// TwinCAT 3 PLC project TcoIo
// Title: TcoIo
// Company: Vortex.Library
// Author: Inxton
// ProjectVersion: 0.6.0.913
// ProgramVersion: 3.1.4023.0
// libraries:
//   Tc2_EtherCAT, * (Beckhoff Automation GmbH)
//   Tc2_Standard, * (Beckhoff Automation GmbH)
//   Tc2_System, * (Beckhoff Automation GmbH)
//   Tc3_Module, * (Beckhoff Automation GmbH)
//   TcoCore, 0.6.0.913 (Vortex.Library)
// project tree:
//   Diagnostics/EtherCAT/MasterDevice/Base/ EtcMasterBase_62654B43.TcDUT, SyncUnitsBase_AD6C35CE.TcDUT, SyncUnitTaskBase_FCD3CBF3.TcDUT, SyncUnitTasksBase_7C8711EB.TcDUT
//   Diagnostics/EtherCAT/MasterDevice/SyncUnit/ InfoData_8649EEEB.TcDUT, ITcoSyncUnit.TcIO, SyncUnitState.TcDUT, SyncUnitTask_AB2F5079.TcDUT, TcoSyncUnit.TcPOU
//   Diagnostics/EtherCAT/SlaveDevice/Base/ EtcSlaveBase_82538BE2.TcDUT, EtcSlaveBoxBase_77A0E4A7.TcDUT, EtcSlaveEndTerminalBase_866C7F0C.TcDUT, EtcSlaveTerminalBase_947E5A46.TcDUT
//   Diagnostics/EtherCAT/MasterDevice/ InfoData_84133AC9.TcDUT, Inputs_A65FACA4.TcDUT, Outputs_23C0ED1D.TcDUT, TcoEthercatDiagnosticsTask.TcPOU, TcoEthercatMasterDeviceState.TcDUT, ITcoEthercatMasterDevice.TcIO, TcoEthercatMasterDevice.TcPOU
//   Diagnostics/EtherCAT/MasterDevice/Messenger/ DiagnosticsMessenger.TcPOU, DiagnosticsMessengers.TcPOU
//   Diagnostics/EtherCAT/SlaveDevice/InfoData/ InfoData_23CBA837.TcDUT, InfoData_6F19DB2B.TcDUT
//   Diagnostics/EtherCAT/SlaveDevice/Inputs/ InputBase_8311D824.TcDUT
//   Diagnostics/EtherCAT/SlaveDevice/Outputs/ OutputBase_10CEE7DE.TcDUT
//   Diagnostics/EtherCAT/SlaveDevice/WcState/ WcState_0B2B16F9.TcDUT, WcState_9091E0EB.TcDUT
//   Diagnostics/EtherCAT/ TcoEthercat.TcGVL
//   Diagnostics/ProfinetComponent/ TcoPnIoComponent.TcPOU
//   EtherCAT/ eEcatState.TcDUT, eLinkState.TcDUT, ITcoEcatComponent.TcIO, TcoEcatSlaveState.TcPOU, TcoEcatComponent.TcPOU
//   / PlcTask.TcTTO
//   POUs/ MAIN.TcPOU
//   SpecialPlcTypes/ TcoAmsAddr.TcDUT, TcoAmsNetId.TcDUT
// real-time tasks:
//   TASK PlcTask: cycle T#15ms, priority 12, ADS port 350
//   TASK PlcTask1: cycle T#15ms, priority 6, ADS port 351
//   TASK PlcTask2: cycle T#10ms, priority 20, ADS port 352
// I/O:
//   DEVICE Device 1 (EtherCAT) (disabled), AmsNetId 172.20.10.110.2.1
//     Term 1 (EK1200) [EK1200-5000 EtherCAT Power supply (2A E-Bus)]
//       Term 2 (EL6002) [EL6002 Interface 2Ch. (RS232)]
//       Term 3 (EL1809) [EL1809 16Ch. Dig. Input 24V, 3ms]
//       Term 4 (EL2809) [EL2809 16Ch. Dig. Output 24V, 0.5A]
//       Term 5 (EL4004) [EL4004 4Ch. Ana. Output 0-10V, 12bit]
//       Term 6 (EL2809) [EL2809 16Ch. Dig. Output 24V, 0.5A]
//       Term 7 (EL6001) [EL6001 Interface (RS232)]
//       Term 8 (EL9011) [EL9011 End Terminal]
//   DEVICE Device 2 (EtherCAT) (disabled), AmsNetId 172.20.10.110.3.1
//     Term 9 (EK1100) [EK1100 EtherCAT Coupler (2A E-Bus)]
//       Term 10 (EK1122) [EK1122 2 port EtherCAT junction]
//         Term 11 (EK1100) [EK1100 EtherCAT Coupler (2A E-Bus)]
//           Term 12 (EL3174-0002) [EL3174-0002 4Ch. Ana. Input +/-10V, +/-20mA 16 Bit, Isolated Channels]
//           Term 13 (EL6001) [EL6001 Interface (RS232)]
//           Term 14 (EL3011) [EL3011 4Ch. Ana. Input 0-20mA DIFF]
//           Term 15 (EL2008) [EL2008 8Ch. Dig. Output 24V, 0.5A]
//           Term 16 (EL2008) [EL2008 8Ch. Dig. Output 24V, 0.5A]
//           Term 17 (EK1110) [EK1110 EtherCAT extension]
//         Term 18 (EK1100) [EK1100 EtherCAT Coupler (2A E-Bus)]
//           Term 19 (EL1809) [EL1809 16Ch. Dig. Input 24V, 3ms]
//           Term 20 (EL2809) [EL2809 16Ch. Dig. Output 24V, 0.5A]
//           Term 21 (EL1809) [EL1809 16Ch. Dig. Input 24V, 3ms]
//           Term 22 (EL3011) [EL3011 4Ch. Ana. Input 0-20mA DIFF]
//           Term 29 (EL9011) [EL9011 End Terminal]
//         Term 23 (EK1100) [EK1100 EtherCAT Coupler (2A E-Bus)]
//           Term 24 (EK1122) [EK1122 2 port EtherCAT junction]
//             Term 25 (EK1100) [EK1100 EtherCAT Coupler (2A E-Bus)]
//               Term 26 (EL1819) [EL1819 16Ch. Dig. Input 24V, 10µs]
//               Term 27 (EL1819) [EL1819 16Ch. Dig. Input 24V, 10µs]
//               Term 30 (EL9011) [EL9011 End Terminal]
//             Term 28 (EK1100) [EK1100 EtherCAT Coupler (2A E-Bus)]
//               Term 29 (EL2788) [EL2788 8Ch. Dig. Output 24V AC/DC, 2A]
//               Term 30 (EL3773) [EL3773 3 Ch. Power Monitoring, Oversample]
//               Term 31 (EL9011) [EL9011 End Terminal]
//           Term 31 (EL3773) [EL3773 3 Ch. Power Monitoring, Oversample]
//           Term 32 (EL2258) [EL2258 8Ch. Dig Output 24V with Multi-Time-Stamp]
//           Term 33 (EL3164) [EL3164 4Ch. Ana. Input 0-10V]
//           Term 32 (EL9011) [EL9011 End Terminal]
//       Term 34 (EL3403) [EL3403 3Ch. Power Measuring]
//       Term 35 (EL6001) [EL6001 Interface (RS232)]
//       Term 36 (EL3024) [EL3024 4Ch. Ana. Input 4-20mA DIFF]
//       Term 33 (EL9011) [EL9011 End Terminal]
//   DEVICE Device 3 (EtherCAT) (disabled), AmsNetId 172.20.10.110.4.1
//     Term 146 (EK1100) [EK1100 EtherCAT Coupler (2A E-Bus)]
//       Term 147 (EK1122) [EK1122 2 port EtherCAT junction]
//         Term 153 (EK1100) [EK1100 EtherCAT Coupler (2A E-Bus)]
//           Term 154 (EK1122) [EK1122 2 port EtherCAT junction]
//             Term 157 (EK1100) [EK1100 EtherCAT Coupler (2A E-Bus)]
//               Term 159 (EL1809) [EL1809 16Ch. Dig. Input 24V, 3ms]
//             Term 158 (EK1100) [EK1100 EtherCAT Coupler (2A E-Bus)]
//               Term 160 (EL1809) [EL1809 16Ch. Dig. Input 24V, 3ms]
//           Term 155 (EL2008) [EL2008 8Ch. Dig. Output 24V, 0.5A]
//           Term 156 (EL2008) [EL2008 8Ch. Dig. Output 24V, 0.5A]
//         Term 178 (EK1100) [EK1100 EtherCAT Coupler (2A E-Bus)]
//           Term 179 (EK1122) [EK1122 2 port EtherCAT junction]
//             Term 180 (EK1100) [EK1100 EtherCAT Coupler (2A E-Bus)]
//               Term 181 (EL1809) [EL1809 16Ch. Dig. Input 24V, 3ms]
//             Term 182 (EK1100) [EK1100 EtherCAT Coupler (2A E-Bus)]
//               Term 183 (EL1809) [EL1809 16Ch. Dig. Input 24V, 3ms]
//           Term 184 (EL2008) [EL2008 8Ch. Dig. Output 24V, 0.5A]
//           Term 185 (EL2008) [EL2008 8Ch. Dig. Output 24V, 0.5A]
//       Term 186 (EK1122) [EK1122 2 port EtherCAT junction]
//         Term 187 (EK1100) [EK1100 EtherCAT Coupler (2A E-Bus)]
//           Term 188 (EK1122) [EK1122 2 port EtherCAT junction]
//             Term 189 (EK1100) [EK1100 EtherCAT Coupler (2A E-Bus)]
//               Term 193 (EL1809) [EL1809 16Ch. Dig. Input 24V, 3ms]
//             Term 194 (EK1100) [EK1100 EtherCAT Coupler (2A E-Bus)]
//               Term 200 (EL1809) [EL1809 16Ch. Dig. Input 24V, 3ms]
//           Term 204 (EL2008) [EL2008 8Ch. Dig. Output 24V, 0.5A]
//           Term 205 (EL2008) [EL2008 8Ch. Dig. Output 24V, 0.5A]
//         Term 207 (EK1100) [EK1100 EtherCAT Coupler (2A E-Bus)]
//           Term 230 (EK1122) [EK1122 2 port EtherCAT junction]
//             Term 231 (EK1100) [EK1100 EtherCAT Coupler (2A E-Bus)]
//               Term 232 (EL1809) [EL1809 16Ch. Dig. Input 24V, 3ms]
//             Term 233 (EK1100) [EK1100 EtherCAT Coupler (2A E-Bus)]
//               Term 234 (EL1809) [EL1809 16Ch. Dig. Input 24V, 3ms]
//           Term 235 (EL2008) [EL2008 8Ch. Dig. Output 24V, 0.5A]
//           Term 236 (EL2008) [EL2008 8Ch. Dig. Output 24V, 0.5A]
//       Term 148 (EL1809) [EL1809 16Ch. Dig. Input 24V, 3ms]
//       Term 149 (EL1809) [EL1809 16Ch. Dig. Input 24V, 3ms]
//       Term 150 (EL1809) [EL1809 16Ch. Dig. Input 24V, 3ms]
//       Term 151 (EL1809) [EL1809 16Ch. Dig. Input 24V, 3ms]
//       Term 152 (EL1809) [EL1809 16Ch. Dig. Input 24V, 3ms]
//       Term 288 (EK1122) [EK1122 2 port EtherCAT junction]
//         Term 289 (EK1100) [EK1100 EtherCAT Coupler (2A E-Bus)]
//           Term 237 (EK1122) [EK1122 2 port EtherCAT junction]
//             Drive 238 (AX5101-0000-0214) [AX5101-0000-0214 EtherCAT Drive (SoE, 1 Ch.)]
//           Term 293 (EL1809) [EL1809 16Ch. Dig. Input 24V, 3ms]
//         Term 294 (EK1100) [EK1100 EtherCAT Coupler (2A E-Bus)]
//           Term 300 (EL1809) [EL1809 16Ch. Dig. Input 24V, 3ms]
//           Term 304 (EL2008) [EL2008 8Ch. Dig. Output 24V, 0.5A]
//           Term 305 (EL2008) [EL2008 8Ch. Dig. Output 24V, 0.5A]
//         Term 307 (EK1100) [EK1100 EtherCAT Coupler (2A E-Bus)]
//           Term 330 (EK1122) [EK1122 2 port EtherCAT junction]
//             Term 331 (EK1100) [EK1100 EtherCAT Coupler (2A E-Bus)]
//               Term 332 (EL1809) [EL1809 16Ch. Dig. Input 24V, 3ms]
//             Term 333 (EK1100) [EK1100 EtherCAT Coupler (2A E-Bus)]
//               Term 334 (EL1809) [EL1809 16Ch. Dig. Input 24V, 3ms]
//           Term 335 (EL2008) [EL2008 8Ch. Dig. Output 24V, 0.5A]
//           Term 336 (EL2008) [EL2008 8Ch. Dig. Output 24V, 0.5A]
//       Term 1158 (EL2008) [EL2008 8Ch. Dig. Output 24V, 0.5A]
//       Term 1159 (EL2008) [EL2008 8Ch. Dig. Output 24V, 0.5A]
//       Term 1160 (EL2008) [EL2008 8Ch. Dig. Output 24V, 0.5A]
//       Term 1161 (EL2008) [EL2008 8Ch. Dig. Output 24V, 0.5A]
//       Term 1162 (EL2008) [EL2008 8Ch. Dig. Output 24V, 0.5A]
//       Term 1163 (EL2008) [EL2008 8Ch. Dig. Output 24V, 0.5A]
//   DEVICE Device 4 (EtherCAT) (disabled), AmsNetId 172.20.10.110.5.1
//     R1 (EK1100) [EK1100 EtherCAT Coupler (2A E-Bus)]
//       R1_A2_EC (EK1122) [EK1122 2 port EtherCAT junction]
//         Servo_A10_1 (AX5106-0000-0203) [AX5106-0000-0203 EtherCAT Drive (SoE, 1 Ch.)]
//         Servo_A10_2 (AX5106-0000-0203) [AX5106-0000-0203 EtherCAT Drive (SoE, 1 Ch.)]
//         Servo_A10_3 (AX5106-0000-0203) [AX5106-0000-0203 EtherCAT Drive (SoE, 1 Ch.)]
//       R1_A3_EC (EK1122) [EK1122 2 port EtherCAT junction]
//         VI-2 (AES-D-BC-ECAT) [AES Fieldbus Coupler]
//           modules: Module 1 (32 Byte Valve Unit (0x7F))
//         VI-4 (AES-D-BC-ECAT) [AES Fieldbus Coupler]
//           modules: Module 1 (32 Byte Valve Unit (0x7F))
//       R1_A4_EC (EK1122) [EK1122 2 port EtherCAT junction]
//         R1_A4_X1 (EK1100) [EK1100 EtherCAT Coupler (2A E-Bus)]
//           R1_A4_X1_PN (EL6631) [EL6631 PROFINET IO Controller]
//           R1_A4_X1_IA1 (EL1809) [EL1809 16Ch. Dig. Input 24V, 3ms]
//           R1_A4_X1_IA2 (EL1809) [EL1809 16Ch. Dig. Input 24V, 3ms]
//           R1_A4_X1_IA3 (EL1809) [EL1809 16Ch. Dig. Input 24V, 3ms]
//           R1_A4_X1_IA4 (EL1809) [EL1809 16Ch. Dig. Input 24V, 3ms]
//           R1_A4_X1_QA1 (EL2809) [EL2809 16Ch. Dig. Output 24V, 0.5A]
//           R1_A4_X1_QA2 (EL2809) [EL2809 16Ch. Dig. Output 24V, 0.5A]
//           R1_A4_X1_QA3 (EL2809) [EL2809 16Ch. Dig. Output 24V, 0.5A]
//           R1_A4_X1_EndTerminal (EL9010) [EL9010 End Terminal]
//         R1_A4_X2 (EK1100) [EK1100 EtherCAT Coupler (2A E-Bus)]
//           R1_A4_X2_A2 (EK1122) [EK1122 2 port EtherCAT junction]
//             R1_A4_X2_A2_VI1 (AES-D-BC-ECAT) [AES Fieldbus Coupler]
//               modules: Module 1 (32 Byte Valve Unit (0x7F))
//             REX_350 (IMecat) [IMecat]
//           R1_A4_X2_IA1 (EL1809) [EL1809 16Ch. Dig. Input 24V, 3ms]
//           R1_A4_X2_IA2 (EL1809) [EL1809 16Ch. Dig. Input 24V, 3ms]
//           R1_A4_X2_IA3 (EL1809) [EL1809 16Ch. Dig. Input 24V, 3ms]
//           R1_A4_X2_IA4 (EL1809) [EL1809 16Ch. Dig. Input 24V, 3ms]
//           R1_A4_X2_IA5 (EL1809) [EL1809 16Ch. Dig. Input 24V, 3ms]
//           R1_A4_X2_QA1 (EL2809) [EL2809 16Ch. Dig. Output 24V, 0.5A]
//           R1_A4_X2_QA2 (EL2809) [EL2809 16Ch. Dig. Output 24V, 0.5A]
//           R1_A4_X2_QA3 (EL2809) [EL2809 16Ch. Dig. Output 24V, 0.5A]
//           R1_A4_X2_EndTerminal (EL9010) [EL9010 End Terminal]
//       R1_A5_DI (EL1809) [EL1809 16Ch. Dig. Input 24V, 3ms]
//       R1_A6_DI (EL1809) [EL1809 16Ch. Dig. Input 24V, 3ms]
//       R1_A7_DI (EL1809) [EL1809 16Ch. Dig. Input 24V, 3ms]
//       R1_A8_DI (EL1809) [EL1809 16Ch. Dig. Input 24V, 3ms]
//       R1_A9_DI (EL1809) [EL1809 16Ch. Dig. Input 24V, 3ms]
//       R1_A10_DI (EL1809) [EL1809 16Ch. Dig. Input 24V, 3ms]
//       R1_A11_DI (EL1809) [EL1809 16Ch. Dig. Input 24V, 3ms]
//       R1_A12_DI (EL1809) [EL1809 16Ch. Dig. Input 24V, 3ms]
//       R1_A13_DI (EL1809) [EL1809 16Ch. Dig. Input 24V, 3ms]
//       R1_A14_DI (EL1809) [EL1809 16Ch. Dig. Input 24V, 3ms]
//       R1_A15_DI (EL1809) [EL1809 16Ch. Dig. Input 24V, 3ms]
//       R1_A16_DI (EL1809) [EL1809 16Ch. Dig. Input 24V, 3ms]
//       R1_A17_DI (EL1809) [EL1809 16Ch. Dig. Input 24V, 3ms]
//       R1_A18_DO (EL2809) [EL2809 16Ch. Dig. Output 24V, 0.5A]
//       R1_A19_DO (EL2809) [EL2809 16Ch. Dig. Output 24V, 0.5A]
//       R1_A20_DO (EL2809) [EL2809 16Ch. Dig. Output 24V, 0.5A]
//       R1_A21_DO (EL2809) [EL2809 16Ch. Dig. Output 24V, 0.5A]
//       R1_A22_DO (EL2809) [EL2809 16Ch. Dig. Output 24V, 0.5A]
//       R1_A23_DO (EL2809) [EL2809 16Ch. Dig. Output 24V, 0.5A]
//       R1_EndTerminal (EL9011) [EL9011 End Terminal]
//     R2 (EK1100) [EK1100 EtherCAT Coupler (2A E-Bus)]
//       R2_A2_EC (EK1122) [EK1122 2 port EtherCAT junction]
//         Servo_A20-2 (AX5103-0000-0203) [AX5103-0000-0203 EtherCAT Drive (SoE, 1 Ch.)]
//         VI-3 (AES-D-BC-ECAT) [AES Fieldbus Coupler]
//           modules: Module 1 (32 Byte Valve Unit (0x7F))
//       R2_A3_DI (EL1809) [EL1809 16Ch. Dig. Input 24V, 3ms]
//       R2_A4_DI (EL1809) [EL1809 16Ch. Dig. Input 24V, 3ms]
//       R2_A5_DI (EL1809) [EL1809 16Ch. Dig. Input 24V, 3ms]
//       R2_A6_DI (EL1809) [EL1809 16Ch. Dig. Input 24V, 3ms]
//       R2_A7_DI (EL1809) [EL1809 16Ch. Dig. Input 24V, 3ms]
//       R2_A8_DI (EL1809) [EL1809 16Ch. Dig. Input 24V, 3ms]
//       R2_A9_DI (EL1809) [EL1809 16Ch. Dig. Input 24V, 3ms]
//       R2_A10_DI (EL1809) [EL1809 16Ch. Dig. Input 24V, 3ms]
//       R2_A11_DC (EL7332) [EL7332 2Ch. DC motor output stage (24V, 1.5A)]
//       R2_A12_DI (EL1809) [EL1809 16Ch. Dig. Input 24V, 3ms]
//       R2_A13_DI (EL1809) [EL1809 16Ch. Dig. Input 24V, 3ms]
//       R2_A14_DI (EL1809) [EL1809 16Ch. Dig. Input 24V, 3ms]
//       R2_A15_DO (EL2809) [EL2809 16Ch. Dig. Output 24V, 0.5A]
//       R2_A16_DO (EL2809) [EL2809 16Ch. Dig. Output 24V, 0.5A]
//       R2_A17_DO (EL2809) [EL2809 16Ch. Dig. Output 24V, 0.5A]
//       R2_A18_DO (EL2809) [EL2809 16Ch. Dig. Output 24V, 0.5A]
//       R2_A19_DO (EL2809) [EL2809 16Ch. Dig. Output 24V, 0.5A]
//       R2_EndTerminal (EL9011) [EL9011 End Terminal]
//     R3 (EK1100) [EK1100 EtherCAT Coupler (2A E-Bus)]
//       R3_A2_EC (EK1122) [EK1122 2 port EtherCAT junction]
//         R3_FESTO (CMMP-AS V4p0 CiA402) [CMMP-AS V4p0 CiA402]
//         VI-1 (AES-D-BC-ECAT) [AES Fieldbus Coupler]
//           modules: Module 1 (32 Byte Valve Unit (0x7F))
//       R3_A3_DI (EL1809) [EL1809 16Ch. Dig. Input 24V, 3ms]
//       R3_A4_DI (EL1809) [EL1809 16Ch. Dig. Input 24V, 3ms]
//       R3_A5_DI (EL1809) [EL1809 16Ch. Dig. Input 24V, 3ms]
//       R3_A6_DI (EL1809) [EL1809 16Ch. Dig. Input 24V, 3ms]
//       R3_A7_DI (EL1809) [EL1809 16Ch. Dig. Input 24V, 3ms]
//       R3_A8_DI (EL1809) [EL1809 16Ch. Dig. Input 24V, 3ms]
//       R3_A9_DO (EL2809) [EL2809 16Ch. Dig. Output 24V, 0.5A]
//       R3_A10_DO (EL2809) [EL2809 16Ch. Dig. Output 24V, 0.5A]
//       R3_EndTerminal (EL9011) [EL9011 End Terminal]
//     R4 (EK1100) [EK1100 EtherCAT Coupler (2A E-Bus)]
//       R4_A2_EC (EK1122) [EK1122 2 port EtherCAT junction]
//         R4_FESTO (CMMP-AS V4p0 CiA402) [CMMP-AS V4p0 CiA402]
//         RH (EK1100) [EK1100 EtherCAT Coupler (2A E-Bus)]
//           RH_A2 (EK1122) [EK1122 2 port EtherCAT junction]
//             RH_SAFETY (Flexi Gateway GETC1) [FLX0-GETC100]
//             RH_A2_X2 (EK1100) [EK1100 EtherCAT Coupler (2A E-Bus)]
//               RH_A2_X2_A2 (EL7211-0010) [EL7211-0010 1Ch. MDP742 Servo motor output stage with OCT (50V, 4.5A RMS)]
//               RH_A2_X2_A3 (EL1809) [EL1809 16Ch. Dig. Input 24V, 3ms]
//               RH_A2_X2_A4 (EL2809) [EL2809 16Ch. Dig. Output 24V, 0.5A]
//               Term 1057 (EL9011) [EL9011 End Terminal]
//           RH_A3 (EL6631) [EL6631 PROFINET IO Controller]
//           RH_A4 (EL1809) [EL1809 16Ch. Dig. Input 24V, 3ms]
//           RH_A5 (EL1809) [EL1809 16Ch. Dig. Input 24V, 3ms]
//           RH_A6 (EL1809) [EL1809 16Ch. Dig. Input 24V, 3ms]
//           RH_A7 (EL2809) [EL2809 16Ch. Dig. Output 24V, 0.5A]
//           RH_A8 (EL1809) [EL1809 16Ch. Dig. Input 24V, 3ms]
//           RH_A9 (EL2809) [EL2809 16Ch. Dig. Output 24V, 0.5A]
//           RH_A10 (EL2809) [EL2809 16Ch. Dig. Output 24V, 0.5A]
//           RH_A11 (EL2809) [EL2809 16Ch. Dig. Output 24V, 0.5A]
//           RH_EndTerminal (EL9011) [EL9011 End Terminal]
//       R4_A3_DI (EL1809) [EL1809 16Ch. Dig. Input 24V, 3ms]
//       R4_A4_DI (EL1809) [EL1809 16Ch. Dig. Input 24V, 3ms]
//       R4_A5_DI (EL1809) [EL1809 16Ch. Dig. Input 24V, 3ms]
//       R4_A6_DI (EL1809) [EL1809 16Ch. Dig. Input 24V, 3ms]
//       R4_A7_DI (EL1809) [EL1809 16Ch. Dig. Input 24V, 3ms]
//       R4_EndTerminal (EL9011) [EL9011 End Terminal]
//     R4A (EK1100) [EK1100 EtherCAT Coupler (2A E-Bus)]
//       A2 (EK1122) [EK1122 2 port EtherCAT junction]
//         VI-7 (AES-D-BC-ECAT) [AES Fieldbus Coupler]
//           modules: Module 1 (32 Byte Valve Unit (0x7F))
//       A3 (EL1809) [EL1809 16Ch. Dig. Input 24V, 3ms]
//       A4 (EL1809) [EL1809 16Ch. Dig. Input 24V, 3ms]
//       A5 (EL1809) [EL1809 16Ch. Dig. Input 24V, 3ms]
//       A6 (EL1809) [EL1809 16Ch. Dig. Input 24V, 3ms]
//       A7 (EL3692) [EL3692 2Ch. resistance measurement terminal]
//       A8 (EL3692) [EL3692 2Ch. resistance measurement terminal]
//       A9 (EL2008) [EL2008 8Ch. Dig. Output 24V, 0.5A]
//       A10 (EL2008) [EL2008 8Ch. Dig. Output 24V, 0.5A]
//       R4A_EndTerminal (EL9011) [EL9011 End Terminal]
//     R5 (EK1100) [EK1100 EtherCAT Coupler (2A E-Bus)]
//       R5_A2_EC (EK1122) [EK1122 2 port EtherCAT junction]
//         VI-5 (AES-D-BC-ECAT) [AES Fieldbus Coupler]
//           modules: Module 1 (32 Byte Valve Unit (0x7F))
//       R5_A3_DI (EL1809) [EL1809 16Ch. Dig. Input 24V, 3ms]
//       R5_A4_DI (EL1809) [EL1809 16Ch. Dig. Input 24V, 3ms]
//       R5_A5_DO (EL2809) [EL2809 16Ch. Dig. Output 24V, 0.5A]
//       R5_A6_DO (EL2809) [EL2809 16Ch. Dig. Output 24V, 0.5A]
//       R5_EndTerminal (EL9011) [EL9011 End Terminal]
//     R6 (EK1100) [EK1100 EtherCAT Coupler (2A E-Bus)]
//       R6_A2_DI (EL1809) [EL1809 16Ch. Dig. Input 24V, 3ms]
//       R6_A3_DI (EL1809) [EL1809 16Ch. Dig. Input 24V, 3ms]
//       R6_A4_DI (EL1809) [EL1809 16Ch. Dig. Input 24V, 3ms]
//       R6_A5_DI (EL1809) [EL1809 16Ch. Dig. Input 24V, 3ms]
//       R6_A6_DI (EL1809) [EL1809 16Ch. Dig. Input 24V, 3ms]
//       R6_A7_DI (EL1809) [EL1809 16Ch. Dig. Input 24V, 3ms]
//       R6_A8_DI (EL1809) [EL1809 16Ch. Dig. Input 24V, 3ms]
//       R6_A9_DI (EL1809) [EL1809 16Ch. Dig. Input 24V, 3ms]
//       R6_A10_DI (EL1809) [EL1809 16Ch. Dig. Input 24V, 3ms]
//       R6_A11_DI (EL1809) [EL1809 16Ch. Dig. Input 24V, 3ms]
//       R6_A12_DI (EL1809) [EL1809 16Ch. Dig. Input 24V, 3ms]
//       R6_A13_DI (EL1809) [EL1809 16Ch. Dig. Input 24V, 3ms]
//       R6_A14_DI (EL1809) [EL1809 16Ch. Dig. Input 24V, 3ms]
//       R6_A15_DO (EL2809) [EL2809 16Ch. Dig. Output 24V, 0.5A]
//       R6_A16_DO (EL2809) [EL2809 16Ch. Dig. Output 24V, 0.5A]
//       R6_A17_DO (EL2809) [EL2809 16Ch. Dig. Output 24V, 0.5A]
//       R6_A18_DO (EL2809) [EL2809 16Ch. Dig. Output 24V, 0.5A]
//       R6_EndTerminal (EL9011) [EL9011 End Terminal]
//     R7 (EK1100) [EK1100 EtherCAT Coupler (2A E-Bus)]
//       R7_A2_EC (EK1122) [EK1122 2 port EtherCAT junction]
//         VI-6 (AES-D-BC-ECAT) [AES Fieldbus Coupler]
//           modules: Module 1 (32 Byte Valve Unit (0x7F))
//       R7_A3_DI (EL1809) [EL1809 16Ch. Dig. Input 24V, 3ms]
//       R7_A4_DI (EL1809) [EL1809 16Ch. Dig. Input 24V, 3ms]
//       R7_A5_DI (EL1809) [EL1809 16Ch. Dig. Input 24V, 3ms]
//       R7_A6_DI (EL1809) [EL1809 16Ch. Dig. Input 24V, 3ms]
//       R7_A7_DI (EL1809) [EL1809 16Ch. Dig. Input 24V, 3ms]
//       R7_A8_DI (EL1809) [EL1809 16Ch. Dig. Input 24V, 3ms]
//       R7_A9_DI (EL1809) [EL1809 16Ch. Dig. Input 24V, 3ms]
//       R7_A10_DI (EL1809) [EL1809 16Ch. Dig. Input 24V, 3ms]
//       R7_A11_DI (EL1809) [EL1809 16Ch. Dig. Input 24V, 3ms]
//       R7_A12_DI (EL1809) [EL1809 16Ch. Dig. Input 24V, 3ms]
//       R7_A13_DI (EL2809) [EL2809 16Ch. Dig. Output 24V, 0.5A]
//       R7_A14_DI (EL2809) [EL2809 16Ch. Dig. Output 24V, 0.5A]
//       R7_EndTerminal (EL9011) [EL9011 End Terminal]
//     R8 (EK1100) [EK1100 EtherCAT Coupler (2A E-Bus)]
//       R8_A2 (EK1122) [EK1122 2 port EtherCAT junction]
//         R8_AB0 (EPP1322-0001) [EPP1322-0001 3 port EtherCAT P gateway]
//           R8_AB24 (EPP1008-0001) [EPP1008-0001 8 Ch. Dig. Input 24V, 3ms, M8]
//           R8_AB23 (EPP1008-0001) [EPP1008-0001 8 Ch. Dig. Input 24V, 3ms, M8]
//           R8_AB22 (EPP1008-0001) [EPP1008-0001 8 Ch. Dig. Input 24V, 3ms, M8]
//           R8_AB21 (EPP1008-0001) [EPP1008-0001 8 Ch. Dig. Input 24V, 3ms, M8]
//           R8_AB20 (EPP1008-0001) [EPP1008-0001 8 Ch. Dig. Input 24V, 3ms, M8]
//           R8_AB19 (EPP1008-0001) [EPP1008-0001 8 Ch. Dig. Input 24V, 3ms, M8]
//           R8_AB18 (EPP1008-0001) [EPP1008-0001 8 Ch. Dig. Input 24V, 3ms, M8]
//           R8_AB17 (EPP1008-0001) [EPP1008-0001 8 Ch. Dig. Input 24V, 3ms, M8]
//           R8_AB16 (EPP1008-0001) [EPP1008-0001 8 Ch. Dig. Input 24V, 3ms, M8]
//           R8_AB15 (EPP1008-0001) [EPP1008-0001 8 Ch. Dig. Input 24V, 3ms, M8]
//           R8_AB14 (EPP1008-0001) [EPP1008-0001 8 Ch. Dig. Input 24V, 3ms, M8]
//           R8_AB13 (EPP1008-0001) [EPP1008-0001 8 Ch. Dig. Input 24V, 3ms, M8]
//           Box 379 (EPP1332-0001) [EPP1332-0001 3 port EtherCAT P junction, power refreshing]
//           R8_AB12 (EPP1008-0001) [EPP1008-0001 8 Ch. Dig. Input 24V, 3ms, M8]
//           R8_AB11 (EPP1008-0001) [EPP1008-0001 8 Ch. Dig. Input 24V, 3ms, M8]
//           R8_AB10 (EPP1008-0001) [EPP1008-0001 8 Ch. Dig. Input 24V, 3ms, M8]
//           R8_AB9 (EPP1008-0001) [EPP1008-0001 8 Ch. Dig. Input 24V, 3ms, M8]
//           R8_AB8 (EPP1008-0001) [EPP1008-0001 8 Ch. Dig. Input 24V, 3ms, M8]
//           R8_AB7 (EPP1008-0001) [EPP1008-0001 8 Ch. Dig. Input 24V, 3ms, M8]
//           R8_AB6 (EPP1008-0001) [EPP1008-0001 8 Ch. Dig. Input 24V, 3ms, M8]
//           R8_AB5 (EPP1008-0001) [EPP1008-0001 8 Ch. Dig. Input 24V, 3ms, M8]
//           R8_AB4 (EPP1008-0001) [EPP1008-0001 8 Ch. Dig. Input 24V, 3ms, M8]
//           R8_AB3 (EPP1008-0001) [EPP1008-0001 8 Ch. Dig. Input 24V, 3ms, M8]
//           R8_AB2 (EPP1008-0001) [EPP1008-0001 8 Ch. Dig. Input 24V, 3ms, M8]
//           R8_AB1 (EPP1008-0001) [EPP1008-0001 8 Ch. Dig. Input 24V, 3ms, M8]
//       R8_A3 (EK1122) [EK1122 2 port EtherCAT junction]
//         VI-10 (AES-D-BC-ECAT) [AES Fieldbus Coupler]
//           modules: Module 1 (32 Byte Valve Unit (0x7F))
//         VI-9 (AES-D-BC-ECAT) [AES Fieldbus Coupler]
//           modules: Module 1 (32 Byte Valve Unit (0x7F))
//       R8_A5 (EL1809) [EL1809 16Ch. Dig. Input 24V, 3ms]
//       R8_A6 (EL2809) [EL2809 16Ch. Dig. Output 24V, 0.5A]
//       R8_A7 (EL2809) [EL2809 16Ch. Dig. Output 24V, 0.5A]
//       R8_A8 (EK1122) [EK1122 2 port EtherCAT junction]
//         RC10_1 (EK1100) [EK1100 EtherCAT Coupler (2A E-Bus)]
//           RC10_A2 (EK1122) [EK1122 2 port EtherCAT junction]
//             RC10_VI (AES-D-BC-ECAT) [AES Fieldbus Coupler]
//               modules: Module 1 (32 Byte Valve Unit (0x7F))
//             RC10_SAFETY (Flexi Soft EtherCAT Gateway) [Flexi Soft EtherCAT Gateway]
//           RC10_A3 (EK1122) [EK1122 2 port EtherCAT junction]
//             RC10_EPP (EPP1322-0001) [EPP1322-0001 3 port EtherCAT P gateway]
//               RC10_AB1 (EPP1008-0001) [EPP1008-0001 8 Ch. Dig. Input 24V, 3ms, M8]
//               RC10_AB2 (EPP1008-0001) [EPP1008-0001 8 Ch. Dig. Input 24V, 3ms, M8]
//               RC10_AB6 (EPP1008-0001) [EPP1008-0001 8 Ch. Dig. Input 24V, 3ms, M8]
//               RC10_AB3 (EPP1008-0001) [EPP1008-0001 8 Ch. Dig. Input 24V, 3ms, M8]
//               RC10_AB4 (EPP1008-0001) [EPP1008-0001 8 Ch. Dig. Input 24V, 3ms, M8]
//               RC10_AB7 (EPP1008-0001) [EPP1008-0001 8 Ch. Dig. Input 24V, 3ms, M8]
//               RC10_AB9 (EPP1008-0001) [EPP1008-0001 8 Ch. Dig. Input 24V, 3ms, M8]
//               RC10_AB10 (EPP1008-0001) [EPP1008-0001 8 Ch. Dig. Input 24V, 3ms, M8]
//               RC10_AB8 (EPP1008-0001) [EPP1008-0001 8 Ch. Dig. Input 24V, 3ms, M8]
//               RC10_AB5 (EPP1008-0001) [EPP1008-0001 8 Ch. Dig. Input 24V, 3ms, M8]
//           RC10_A5 (EL1809) [EL1809 16Ch. Dig. Input 24V, 3ms]
//           RC10_A6 (EL1809) [EL1809 16Ch. Dig. Input 24V, 3ms]
//           RC10_A7 (EL2809) [EL2809 16Ch. Dig. Output 24V, 0.5A]
//           RC10_A8 (EL2809) [EL2809 16Ch. Dig. Output 24V, 0.5A]
//           RC10_A9 (EL2809) [EL2809 16Ch. Dig. Output 24V, 0.5A]
//           RC10_1_EndTerminal (EL9011) [EL9011 End Terminal]
//         RC10_2 (EK1100) [EK1100 EtherCAT Coupler (2A E-Bus)]
//           RC10_B1 (EL7041-1000) [EL7041-1000 1Ch. Stepper motor output stage (50V, 5A, standard)]
//           RC10_B2 (EL7041-1000) [EL7041-1000 1Ch. Stepper motor output stage (50V, 5A, standard)]
//           RC10_C11 (EL7041-1000) [EL7041-1000 1Ch. Stepper motor output stage (50V, 5A, standard)]
//           RC10_C12 (EL7041-1000) [EL7041-1000 1Ch. Stepper motor output stage (50V, 5A, standard)]
//           RC10_C21 (EL7041-1000) [EL7041-1000 1Ch. Stepper motor output stage (50V, 5A, standard)]
//           RC10_C22 (EL7041-1000) [EL7041-1000 1Ch. Stepper motor output stage (50V, 5A, standard)]
//           RC10_2_EndTerminal (EL9010) [EL9010 End Terminal]
//         RC20_1 (EK1100) [EK1100 EtherCAT Coupler (2A E-Bus)]
//           RC20_A2 (EK1122) [EK1122 2 port EtherCAT junction]
//             RC20_VI (AES-D-BC-ECAT) [AES Fieldbus Coupler]
//               modules: Module 1 (32 Byte Valve Unit (0x7F))
//             RC20_SAFETY (Flexi Soft EtherCAT Gateway) [Flexi Soft EtherCAT Gateway]
//           RC20_A3 (EK1122) [EK1122 2 port EtherCAT junction]
//             RC20_EPP (EPP1322-0001) [EPP1322-0001 3 port EtherCAT P gateway]
//               RC20_AB1 (EPP1008-0001) [EPP1008-0001 8 Ch. Dig. Input 24V, 3ms, M8]
//               RC20_AB2 (EPP1008-0001) [EPP1008-0001 8 Ch. Dig. Input 24V, 3ms, M8]
//               RC20_AB6 (EPP1008-0001) [EPP1008-0001 8 Ch. Dig. Input 24V, 3ms, M8]
//               RC20_AB3 (EPP1008-0001) [EPP1008-0001 8 Ch. Dig. Input 24V, 3ms, M8]
//               RC20_AB4 (EPP1008-0001) [EPP1008-0001 8 Ch. Dig. Input 24V, 3ms, M8]
//               RC20_AB7 (EPP1008-0001) [EPP1008-0001 8 Ch. Dig. Input 24V, 3ms, M8]
//               RC20_AB9 (EPP1008-0001) [EPP1008-0001 8 Ch. Dig. Input 24V, 3ms, M8]
//               RC20_AB10 (EPP1008-0001) [EPP1008-0001 8 Ch. Dig. Input 24V, 3ms, M8]
//               RC20_AB8 (EPP1008-0001) [EPP1008-0001 8 Ch. Dig. Input 24V, 3ms, M8]
//               RC20_AB5 (EPP1008-0001) [EPP1008-0001 8 Ch. Dig. Input 24V, 3ms, M8]
//           RC20_A5 (EL1809) [EL1809 16Ch. Dig. Input 24V, 3ms]
//           RC20_A6 (EL1809) [EL1809 16Ch. Dig. Input 24V, 3ms]
//           RC20_A7 (EL2809) [EL2809 16Ch. Dig. Output 24V, 0.5A]
//           RC20_A8 (EL2809) [EL2809 16Ch. Dig. Output 24V, 0.5A]
//           RC20_A9 (EL2809) [EL2809 16Ch. Dig. Output 24V, 0.5A]
//           RC20_1_EndTerminal (EL9010) [EL9010 End Terminal]
//         RC20_2 (EK1100) [EK1100 EtherCAT Coupler (2A E-Bus)]
//           RC20_B1 (EL7041-1000) [EL7041-1000 1Ch. Stepper motor output stage (50V, 5A, standard)]
//           RC20_B2 (EL7041-1000) [EL7041-1000 1Ch. Stepper motor output stage (50V, 5A, standard)]
//           RC20_C11 (EL7041-1000) [EL7041-1000 1Ch. Stepper motor output stage (50V, 5A, standard)]
//           RC20_C12 (EL7041-1000) [EL7041-1000 1Ch. Stepper motor output stage (50V, 5A, standard)]
//           RC20_C21 (EL7041-1000) [EL7041-1000 1Ch. Stepper motor output stage (50V, 5A, standard)]
//           RC20_C22 (EL7041-1000) [EL7041-1000 1Ch. Stepper motor output stage (50V, 5A, standard)]
//           RC20_2_EndTerminal (EL9010) [EL9010 End Terminal]
//       R8_A9 (EK1122) [EK1122 2 port EtherCAT junction]
//         RC30_1 (EK1100) [EK1100 EtherCAT Coupler (2A E-Bus)]
//           RC30_A2 (EK1122) [EK1122 2 port EtherCAT junction]
//             RC30_VI (AES-D-BC-ECAT) [AES Fieldbus Coupler]
//               modules: Module 1 (32 Byte Valve Unit (0x7F))
//             RC30_SAFETY (Flexi Soft EtherCAT Gateway) [Flexi Soft EtherCAT Gateway]
//           RC30_A3 (EK1122) [EK1122 2 port EtherCAT junction]
//             RC30_EPP (EPP1322-0001) [EPP1322-0001 3 port EtherCAT P gateway]
//               RC30_AB1 (EPP1008-0001) [EPP1008-0001 8 Ch. Dig. Input 24V, 3ms, M8]
//               RC30_AB2 (EPP1008-0001) [EPP1008-0001 8 Ch. Dig. Input 24V, 3ms, M8]
//               RC30_AB6 (EPP1008-0001) [EPP1008-0001 8 Ch. Dig. Input 24V, 3ms, M8]
//               RC30_AB3 (EPP1008-0001) [EPP1008-0001 8 Ch. Dig. Input 24V, 3ms, M8]
//               RC30_AB4 (EPP1008-0001) [EPP1008-0001 8 Ch. Dig. Input 24V, 3ms, M8]
//               RC30_AB7 (EPP1008-0001) [EPP1008-0001 8 Ch. Dig. Input 24V, 3ms, M8]
//               RC30_AB9 (EPP1008-0001) [EPP1008-0001 8 Ch. Dig. Input 24V, 3ms, M8]
//               RC30_AB10 (EPP1008-0001) [EPP1008-0001 8 Ch. Dig. Input 24V, 3ms, M8]
//               RC30_AB8 (EPP1008-0001) [EPP1008-0001 8 Ch. Dig. Input 24V, 3ms, M8]
//               RC30_AB5 (EPP1008-0001) [EPP1008-0001 8 Ch. Dig. Input 24V, 3ms, M8]
//           RC30_A5 (EL1809) [EL1809 16Ch. Dig. Input 24V, 3ms]
//           RC30_A6 (EL1809) [EL1809 16Ch. Dig. Input 24V, 3ms]
//           RC30_A7 (EL2809) [EL2809 16Ch. Dig. Output 24V, 0.5A]
//           RC30_A8 (EL2809) [EL2809 16Ch. Dig. Output 24V, 0.5A]
//           RC30_A9 (EL2809) [EL2809 16Ch. Dig. Output 24V, 0.5A]
//           RC30_1_EndTerminal (EL9010) [EL9010 End Terminal]
//         RC30_2 (EK1100) [EK1100 EtherCAT Coupler (2A E-Bus)]
//           RC30_B1 (EL7041-1000) [EL7041-1000 1Ch. Stepper motor output stage (50V, 5A, standard)]
//           RC30_B2 (EL7041-1000) [EL7041-1000 1Ch. Stepper motor output stage (50V, 5A, standard)]
//           RC30_C11 (EL7041-1000) [EL7041-1000 1Ch. Stepper motor output stage (50V, 5A, standard)]
//           RC30_C12 (EL7041-1000) [EL7041-1000 1Ch. Stepper motor output stage (50V, 5A, standard)]
//           RC30_C21 (EL7041-1000) [EL7041-1000 1Ch. Stepper motor output stage (50V, 5A, standard)]
//           RC30_C22 (EL7041-1000) [EL7041-1000 1Ch. Stepper motor output stage (50V, 5A, standard)]
//           RC30_2_EndTerminal (EL9010) [EL9010 End Terminal]
//         RC40_1 (EK1100) [EK1100 EtherCAT Coupler (2A E-Bus)]
//           RC40_A2 (EK1122) [EK1122 2 port EtherCAT junction]
//             RC40_VI (AES-D-BC-ECAT) [AES Fieldbus Coupler]
//               modules: Module 1 (32 Byte Valve Unit (0x7F))
//             RC40_SAFETY (Flexi Soft EtherCAT Gateway) [Flexi Soft EtherCAT Gateway]
//           RC40_A3 (EK1122) [EK1122 2 port EtherCAT junction]
//             RC40_EPP (EPP1322-0001) [EPP1322-0001 3 port EtherCAT P gateway]
//               RC40_AB1 (EPP1008-0001) [EPP1008-0001 8 Ch. Dig. Input 24V, 3ms, M8]
//               RC40_AB2 (EPP1008-0001) [EPP1008-0001 8 Ch. Dig. Input 24V, 3ms, M8]
//               RC40_AB6 (EPP1008-0001) [EPP1008-0001 8 Ch. Dig. Input 24V, 3ms, M8]
//               RC40_AB3 (EPP1008-0001) [EPP1008-0001 8 Ch. Dig. Input 24V, 3ms, M8]
//               RC40_AB4 (EPP1008-0001) [EPP1008-0001 8 Ch. Dig. Input 24V, 3ms, M8]
//               RC40_AB7 (EPP1008-0001) [EPP1008-0001 8 Ch. Dig. Input 24V, 3ms, M8]
//               RC40_AB9 (EPP1008-0001) [EPP1008-0001 8 Ch. Dig. Input 24V, 3ms, M8]
//               RC40_AB10 (EPP1008-0001) [EPP1008-0001 8 Ch. Dig. Input 24V, 3ms, M8]
//               RC40_AB8 (EPP1008-0001) [EPP1008-0001 8 Ch. Dig. Input 24V, 3ms, M8]
//               RC40_AB5 (EPP1008-0001) [EPP1008-0001 8 Ch. Dig. Input 24V, 3ms, M8]
//           RC40_A5 (EL1809) [EL1809 16Ch. Dig. Input 24V, 3ms]
//           RC40_A6 (EL1809) [EL1809 16Ch. Dig. Input 24V, 3ms]
//           RC40_A7 (EL2809) [EL2809 16Ch. Dig. Output 24V, 0.5A]
//           RC40_A8 (EL2809) [EL2809 16Ch. Dig. Output 24V, 0.5A]
//           RC40_A9 (EL2809) [EL2809 16Ch. Dig. Output 24V, 0.5A]
//           RC40_1_EndTerminal (EL9010) [EL9010 End Terminal]
//         RC40_2 (EK1100) [EK1100 EtherCAT Coupler (2A E-Bus)]
//           RC40_B1 (EL7041-1000) [EL7041-1000 1Ch. Stepper motor output stage (50V, 5A, standard)]
//           RC40_B2 (EL7041-1000) [EL7041-1000 1Ch. Stepper motor output stage (50V, 5A, standard)]
//           RC40_C11 (EL7041-1000) [EL7041-1000 1Ch. Stepper motor output stage (50V, 5A, standard)]
//           RC40_C12 (EL7041-1000) [EL7041-1000 1Ch. Stepper motor output stage (50V, 5A, standard)]
//           RC40_C21 (EL7041-1000) [EL7041-1000 1Ch. Stepper motor output stage (50V, 5A, standard)]
//           RC40_C22 (EL7041-1000) [EL7041-1000 1Ch. Stepper motor output stage (50V, 5A, standard)]
//           RC40_2_EndTerminal (EL9010) [EL9010 End Terminal]
//       R8_A10 (EK1122) [EK1122 2 port EtherCAT junction]
//         RC50_1 (EK1100) [EK1100 EtherCAT Coupler (2A E-Bus)]
//           RC50_A2 (EK1122) [EK1122 2 port EtherCAT junction]
//             RC50_VI (AES-D-BC-ECAT) [AES Fieldbus Coupler]
//               modules: Module 1 (32 Byte Valve Unit (0x7F))
//             RC50_SAFETY (Flexi Soft EtherCAT Gateway) [Flexi Soft EtherCAT Gateway]
//           RC50_A3 (EK1122) [EK1122 2 port EtherCAT junction]
//             RC50_EPP (EPP1322-0001) [EPP1322-0001 3 port EtherCAT P gateway]
//               RC50_AB1 (EPP1008-0001) [EPP1008-0001 8 Ch. Dig. Input 24V, 3ms, M8]
//               RC50_AB2 (EPP1008-0001) [EPP1008-0001 8 Ch. Dig. Input 24V, 3ms, M8]
//               RC50_AB6 (EPP1008-0001) [EPP1008-0001 8 Ch. Dig. Input 24V, 3ms, M8]
//               RC50_AB3 (EPP1008-0001) [EPP1008-0001 8 Ch. Dig. Input 24V, 3ms, M8]
//               RC50_AB4 (EPP1008-0001) [EPP1008-0001 8 Ch. Dig. Input 24V, 3ms, M8]
//               RC50_AB7 (EPP1008-0001) [EPP1008-0001 8 Ch. Dig. Input 24V, 3ms, M8]
//               RC50_AB9 (EPP1008-0001) [EPP1008-0001 8 Ch. Dig. Input 24V, 3ms, M8]
//               RC50_AB10 (EPP1008-0001) [EPP1008-0001 8 Ch. Dig. Input 24V, 3ms, M8]
//               RC50_AB8 (EPP1008-0001) [EPP1008-0001 8 Ch. Dig. Input 24V, 3ms, M8]
//               RC50_AB5 (EPP1008-0001) [EPP1008-0001 8 Ch. Dig. Input 24V, 3ms, M8]
//           RC50_A5 (EL1809) [EL1809 16Ch. Dig. Input 24V, 3ms]
//           RC50_A6 (EL1809) [EL1809 16Ch. Dig. Input 24V, 3ms]
//           RC50_A7 (EL2809) [EL2809 16Ch. Dig. Output 24V, 0.5A]
//           RC50_A8 (EL2809) [EL2809 16Ch. Dig. Output 24V, 0.5A]
//           RC50_A9 (EL2809) [EL2809 16Ch. Dig. Output 24V, 0.5A]
//           RC50_1_EndTerminal (EL9010) [EL9010 End Terminal]
//         RC50_2 (EK1100) [EK1100 EtherCAT Coupler (2A E-Bus)]
//           RC50_B1 (EL7041-1000) [EL7041-1000 1Ch. Stepper motor output stage (50V, 5A, standard)]
//           RC50_B2 (EL7041-1000) [EL7041-1000 1Ch. Stepper motor output stage (50V, 5A, standard)]
//           RC50_C11 (EL7041-1000) [EL7041-1000 1Ch. Stepper motor output stage (50V, 5A, standard)]
//           RC50_C12 (EL7041-1000) [EL7041-1000 1Ch. Stepper motor output stage (50V, 5A, standard)]
//           RC50_C21 (EL7041-1000) [EL7041-1000 1Ch. Stepper motor output stage (50V, 5A, standard)]
//           RC50_C22 (EL7041-1000) [EL7041-1000 1Ch. Stepper motor output stage (50V, 5A, standard)]
//           RC50_2_EndTerminal (EL9010) [EL9010 End Terminal]
//         RC60_1 (EK1100) [EK1100 EtherCAT Coupler (2A E-Bus)]
//           RC60_A2 (EK1122) [EK1122 2 port EtherCAT junction]
//             RC60_VI (AES-D-BC-ECAT) [AES Fieldbus Coupler]
//               modules: Module 1 (32 Byte Valve Unit (0x7F))
//             RC60_SAFETY (Flexi Soft EtherCAT Gateway) [Flexi Soft EtherCAT Gateway]
//           RC60_A3 (EK1122) [EK1122 2 port EtherCAT junction]
//             RC60_EPP (EPP1322-0001) [EPP1322-0001 3 port EtherCAT P gateway]
//               RC60_AB1 (EPP1008-0001) [EPP1008-0001 8 Ch. Dig. Input 24V, 3ms, M8]
//               RC60_AB2 (EPP1008-0001) [EPP1008-0001 8 Ch. Dig. Input 24V, 3ms, M8]
//               RC60_AB6 (EPP1008-0001) [EPP1008-0001 8 Ch. Dig. Input 24V, 3ms, M8]
//               RC60_AB3 (EPP1008-0001) [EPP1008-0001 8 Ch. Dig. Input 24V, 3ms, M8]
//               RC60_AB4 (EPP1008-0001) [EPP1008-0001 8 Ch. Dig. Input 24V, 3ms, M8]
//               RC60_AB7 (EPP1008-0001) [EPP1008-0001 8 Ch. Dig. Input 24V, 3ms, M8]
//               RC60_AB9 (EPP1008-0001) [EPP1008-0001 8 Ch. Dig. Input 24V, 3ms, M8]
//               RC60_AB10 (EPP1008-0001) [EPP1008-0001 8 Ch. Dig. Input 24V, 3ms, M8]
//               RC60_AB8 (EPP1008-0001) [EPP1008-0001 8 Ch. Dig. Input 24V, 3ms, M8]
//               RC60_AB5 (EPP1008-0001) [EPP1008-0001 8 Ch. Dig. Input 24V, 3ms, M8]
//           RC60_A5 (EL1809) [EL1809 16Ch. Dig. Input 24V, 3ms]
//           RC60_A6 (EL1809) [EL1809 16Ch. Dig. Input 24V, 3ms]
//           RC60_A7 (EL2809) [EL2809 16Ch. Dig. Output 24V, 0.5A]
//           RC60_A8 (EL2809) [EL2809 16Ch. Dig. Output 24V, 0.5A]
//           RC60_A9 (EL2809) [EL2809 16Ch. Dig. Output 24V, 0.5A]
//           RC60_1_EndTerminal (EL9010) [EL9010 End Terminal]
//         RC60_2 (EK1100) [EK1100 EtherCAT Coupler (2A E-Bus)]
//           RC60_B1 (EL7041-1000) [EL7041-1000 1Ch. Stepper motor output stage (50V, 5A, standard)]
//           RC60_B2 (EL7041-1000) [EL7041-1000 1Ch. Stepper motor output stage (50V, 5A, standard)]
//           RC60_C11 (EL7041-1000) [EL7041-1000 1Ch. Stepper motor output stage (50V, 5A, standard)]
//           RC60_C12 (EL7041-1000) [EL7041-1000 1Ch. Stepper motor output stage (50V, 5A, standard)]
//           RC60_C21 (EL7041-1000) [EL7041-1000 1Ch. Stepper motor output stage (50V, 5A, standard)]
//           RC60_C22 (EL7041-1000) [EL7041-1000 1Ch. Stepper motor output stage (50V, 5A, standard)]
//           RC60_2_EndTerminal (EL9010) [EL9010 End Terminal]
//       R8_A11 (EK1122) [EK1122 2 port EtherCAT junction]
//         RC70_1 (EK1100) [EK1100 EtherCAT Coupler (2A E-Bus)]
//           RC70_A2 (EK1122) [EK1122 2 port EtherCAT junction]
//             RC70_VI (AES-D-BC-ECAT) [AES Fieldbus Coupler]
//               modules: Module 1 (32 Byte Valve Unit (0x7F))
//             RC70_SAFETY (Flexi Soft EtherCAT Gateway) [Flexi Soft EtherCAT Gateway]
//           RC70_A3 (EK1122) [EK1122 2 port EtherCAT junction]
//             RC70_EPP (EPP1322-0001) [EPP1322-0001 3 port EtherCAT P gateway]
//               RC70_AB1 (EPP1008-0001) [EPP1008-0001 8 Ch. Dig. Input 24V, 3ms, M8]
//               RC70_AB2 (EPP1008-0001) [EPP1008-0001 8 Ch. Dig. Input 24V, 3ms, M8]
//               RC70_AB6 (EPP1008-0001) [EPP1008-0001 8 Ch. Dig. Input 24V, 3ms, M8]
//               RC70_AB3 (EPP1008-0001) [EPP1008-0001 8 Ch. Dig. Input 24V, 3ms, M8]
//               RC70_AB4 (EPP1008-0001) [EPP1008-0001 8 Ch. Dig. Input 24V, 3ms, M8]
//               RC70_AB7 (EPP1008-0001) [EPP1008-0001 8 Ch. Dig. Input 24V, 3ms, M8]
//               RC70_AB9 (EPP1008-0001) [EPP1008-0001 8 Ch. Dig. Input 24V, 3ms, M8]
//               RC70_AB10 (EPP1008-0001) [EPP1008-0001 8 Ch. Dig. Input 24V, 3ms, M8]
//               RC70_AB8 (EPP1008-0001) [EPP1008-0001 8 Ch. Dig. Input 24V, 3ms, M8]
//               RC70_AB5 (EPP1008-0001) [EPP1008-0001 8 Ch. Dig. Input 24V, 3ms, M8]
//           RC70_A5 (EL1809) [EL1809 16Ch. Dig. Input 24V, 3ms]
//           RC70_A6 (EL1809) [EL1809 16Ch. Dig. Input 24V, 3ms]
//           RC70_A7 (EL2809) [EL2809 16Ch. Dig. Output 24V, 0.5A]
//           RC70_A8 (EL2809) [EL2809 16Ch. Dig. Output 24V, 0.5A]
//           RC70_A9 (EL2809) [EL2809 16Ch. Dig. Output 24V, 0.5A]
//           RC70_1_EndTerminal (EL9010) [EL9010 End Terminal]
//         RC70_2 (EK1100) [EK1100 EtherCAT Coupler (2A E-Bus)]
//           RC70_B1 (EL7041-1000) [EL7041-1000 1Ch. Stepper motor output stage (50V, 5A, standard)]
//           RC70_B2 (EL7041-1000) [EL7041-1000 1Ch. Stepper motor output stage (50V, 5A, standard)]
//           RC70_C11 (EL7041-1000) [EL7041-1000 1Ch. Stepper motor output stage (50V, 5A, standard)]
//           RC70_C12 (EL7041-1000) [EL7041-1000 1Ch. Stepper motor output stage (50V, 5A, standard)]
//           RC70_C21 (EL7041-1000) [EL7041-1000 1Ch. Stepper motor output stage (50V, 5A, standard)]
//           RC70_C22 (EL7041-1000) [EL7041-1000 1Ch. Stepper motor output stage (50V, 5A, standard)]
//           RC70_2_EndTerminal (EL9010) [EL9010 End Terminal]
//         RC80_1 (EK1100) [EK1100 EtherCAT Coupler (2A E-Bus)] (disabled)
//           RC80_A2 (EK1122) [EK1122 2 port EtherCAT junction]
//             RC80_VI (AES-D-BC-ECAT) [AES Fieldbus Coupler]
//               modules: Module 1 (32 Byte Valve Unit (0x7F))
//             RC80_SAFETY (Flexi Soft EtherCAT Gateway) [Flexi Soft EtherCAT Gateway]
//           RC80_A3 (EK1122) [EK1122 2 port EtherCAT junction]
//             RC80_EPP (EPP1322-0001) [EPP1322-0001 3 port EtherCAT P gateway]
//               RC80_AB1 (EPP1008-0001) [EPP1008-0001 8 Ch. Dig. Input 24V, 3ms, M8]
//               RC80_AB2 (EPP1008-0001) [EPP1008-0001 8 Ch. Dig. Input 24V, 3ms, M8]
//               RC80_AB6 (EPP1008-0001) [EPP1008-0001 8 Ch. Dig. Input 24V, 3ms, M8]
//               RC80_AB3 (EPP1008-0001) [EPP1008-0001 8 Ch. Dig. Input 24V, 3ms, M8]
//               RC80_AB4 (EPP1008-0001) [EPP1008-0001 8 Ch. Dig. Input 24V, 3ms, M8]
//               RC80_AB7 (EPP1008-0001) [EPP1008-0001 8 Ch. Dig. Input 24V, 3ms, M8]
//               RC80_AB9 (EPP1008-0001) [EPP1008-0001 8 Ch. Dig. Input 24V, 3ms, M8]
//               RC80_AB10 (EPP1008-0001) [EPP1008-0001 8 Ch. Dig. Input 24V, 3ms, M8]
//               RC80_AB8 (EPP1008-0001) [EPP1008-0001 8 Ch. Dig. Input 24V, 3ms, M8]
//               RC80_AB5 (EPP1008-0001) [EPP1008-0001 8 Ch. Dig. Input 24V, 3ms, M8]
//           RC80_A5 (EL1809) [EL1809 16Ch. Dig. Input 24V, 3ms]
//           RC80_A6 (EL1809) [EL1809 16Ch. Dig. Input 24V, 3ms]
//           RC80_A7 (EL2809) [EL2809 16Ch. Dig. Output 24V, 0.5A]
//           RC80_A8 (EL2809) [EL2809 16Ch. Dig. Output 24V, 0.5A]
//           RC80_A9 (EL2809) [EL2809 16Ch. Dig. Output 24V, 0.5A]
//           Term 796 (EL9010) [EL9010 End Terminal]
//         RC80_2 (EK1100) [EK1100 EtherCAT Coupler (2A E-Bus)] (disabled)
//           RC80_B1 (EL7041-1000) [EL7041-1000 1Ch. Stepper motor output stage (50V, 5A, standard)]
//           RC80_B2 (EL7041-1000) [EL7041-1000 1Ch. Stepper motor output stage (50V, 5A, standard)]
//           RC80_C11 (EL7041-1000) [EL7041-1000 1Ch. Stepper motor output stage (50V, 5A, standard)]
//           RC80_C12 (EL7041-1000) [EL7041-1000 1Ch. Stepper motor output stage (50V, 5A, standard)]
//           RC80_C21 (EL7041-1000) [EL7041-1000 1Ch. Stepper motor output stage (50V, 5A, standard)]
//           RC80_C22 (EL7041-1000) [EL7041-1000 1Ch. Stepper motor output stage (50V, 5A, standard)]
//           Term 804 (EL9010) [EL9010 End Terminal]
//       R8_A12 (EK1122) [EK1122 2 port EtherCAT junction]
//         RP10 (EK1100) [EK1100 EtherCAT Coupler (2A E-Bus)]
//           RP10_A2 (EK1122) [EK1122 2 port EtherCAT junction]
//             RP10-VI (AES-D-BC-ECAT) [AES Fieldbus Coupler]
//               modules: Module 1 (32 Byte Valve Unit (0x7F))
//             RP10-SAFETY (Flexi Soft EtherCAT Gateway) [Flexi Soft EtherCAT Gateway]
//             RP10-AB0 (EPP1322-0001) [EPP1322-0001 3 port EtherCAT P gateway]
//             RP10-AB1 (EPP1008-0001) [EPP1008-0001 8 Ch. Dig. Input 24V, 3ms, M8]
//             RP10-AB2 (EPP1008-0001) [EPP1008-0001 8 Ch. Dig. Input 24V, 3ms, M8]
//             RP10-AB3 (EPP1008-0001) [EPP1008-0001 8 Ch. Dig. Input 24V, 3ms, M8]
//             RP10-AB4 (EPP1008-0001) [EPP1008-0001 8 Ch. Dig. Input 24V, 3ms, M8]
//           RP10_A4 (EL7041-1000) [EL7041-1000 1Ch. Stepper motor output stage (50V, 5A, standard)]
//           RP10_A5 (EL7041-1000) [EL7041-1000 1Ch. Stepper motor output stage (50V, 5A, standard)]
//           RP10_A6 (EL1809) [EL1809 16Ch. Dig. Input 24V, 3ms]
//           RP10_A7 (EL2809) [EL2809 16Ch. Dig. Output 24V, 0.5A]
//           RP10_EndTerminal (EL9011) [EL9011 End Terminal]
//         RP20 (EK1100) [EK1100 EtherCAT Coupler (2A E-Bus)]
//           RP20_A2 (EK1122) [EK1122 2 port EtherCAT junction]
//             RP20-VI (AES-D-BC-ECAT) [AES Fieldbus Coupler]
//               modules: Module 1 (32 Byte Valve Unit (0x7F))
//             RP20-SAFETY (Flexi Soft EtherCAT Gateway) [Flexi Soft EtherCAT Gateway]
//             RP20-AB0 (EPP1322-0001) [EPP1322-0001 3 port EtherCAT P gateway]
//             RP20-AB1 (EPP1008-0001) [EPP1008-0001 8 Ch. Dig. Input 24V, 3ms, M8]
//             RP20-AB2 (EPP1008-0001) [EPP1008-0001 8 Ch. Dig. Input 24V, 3ms, M8]
//             RP20-AB3 (EPP1008-0001) [EPP1008-0001 8 Ch. Dig. Input 24V, 3ms, M8]
//             RP20-AB4 (EPP1008-0001) [EPP1008-0001 8 Ch. Dig. Input 24V, 3ms, M8]
//           RP20_A4 (EL7041-1000) [EL7041-1000 1Ch. Stepper motor output stage (50V, 5A, standard)]
//           RP20_A5 (EL7041-1000) [EL7041-1000 1Ch. Stepper motor output stage (50V, 5A, standard)]
//           RP20_A6 (EL1809) [EL1809 16Ch. Dig. Input 24V, 3ms]
//           RP20_A7 (EL2809) [EL2809 16Ch. Dig. Output 24V, 0.5A]
//           RP20_EndTerminal (EL9011) [EL9011 End Terminal]
//       R8_A13 (EK1122) [EK1122 2 port EtherCAT junction]
//         RP30 (EK1100) [EK1100 EtherCAT Coupler (2A E-Bus)]
//           RP30_A2 (EK1122) [EK1122 2 port EtherCAT junction]
//             RP30-VI (AES-D-BC-ECAT) [AES Fieldbus Coupler]
//               modules: Module 1 (32 Byte Valve Unit (0x7F))
//             RP30-SAFETY (Flexi Soft EtherCAT Gateway) [Flexi Soft EtherCAT Gateway]
//             RP30-AB0 (EPP1322-0001) [EPP1322-0001 3 port EtherCAT P gateway]
//             RP30-AB1 (EPP1008-0001) [EPP1008-0001 8 Ch. Dig. Input 24V, 3ms, M8]
//             RP30-AB2 (EPP1008-0001) [EPP1008-0001 8 Ch. Dig. Input 24V, 3ms, M8]
//             RP30-AB3 (EPP1008-0001) [EPP1008-0001 8 Ch. Dig. Input 24V, 3ms, M8]
//             RP30-AB4 (EPP1008-0001) [EPP1008-0001 8 Ch. Dig. Input 24V, 3ms, M8]
//           RP30_A4 (EL7041-1000) [EL7041-1000 1Ch. Stepper motor output stage (50V, 5A, standard)]
//           RP30_A5 (EL7041-1000) [EL7041-1000 1Ch. Stepper motor output stage (50V, 5A, standard)]
//           RP30_A6 (EL1809) [EL1809 16Ch. Dig. Input 24V, 3ms]
//           RP30_A7 (EL2809) [EL2809 16Ch. Dig. Output 24V, 0.5A]
//           RP30_EndTerminal (EL9010) [EL9010 End Terminal]
//       R8_Endterminal (EL9010) [EL9010 End Terminal]
//     R9 (EK1100) [EK1100 EtherCAT Coupler (2A E-Bus)]
//       R9_A2 (EK1122) [EK1122 2 port EtherCAT junction]
//         R9_AB0 (EPP1322-0001) [EPP1322-0001 3 port EtherCAT P gateway]
//           R9_AB1 (EPP1008-0001) [EPP1008-0001 8 Ch. Dig. Input 24V, 3ms, M8]
//           R9_AB2 (EPP1008-0001) [EPP1008-0001 8 Ch. Dig. Input 24V, 3ms, M8]
//           R9_AB3 (EPP1008-0001) [EPP1008-0001 8 Ch. Dig. Input 24V, 3ms, M8]
//           R9_AB4 (EPP1008-0001) [EPP1008-0001 8 Ch. Dig. Input 24V, 3ms, M8]
//         R9_SAFETY (Flexi Soft EtherCAT Gateway) [Flexi Soft EtherCAT Gateway]
//       R9_A3 (EK1122) [EK1122 2 port EtherCAT junction]
//         R9_SERVO (IndraDrive MPB20) [IndraDrive MPB20]
//       R9_A5 (EL1809) [EL1809 16Ch. Dig. Input 24V, 3ms]
//       R9_A6 (EL2809) [EL2809 16Ch. Dig. Output 24V, 0.5A]
//       R9_A7 (EL2809) [EL2809 16Ch. Dig. Output 24V, 0.5A]
//       R9_EndTerminal (EL9011) [EL9011 End Terminal]
//     R10 (EK1100) [EK1100 EtherCAT Coupler (2A E-Bus)]
//       R10_A2 (EK1122) [EK1122 2 port EtherCAT junction]
//         R10-VI11 (AES-D-BC-ECAT) [AES Fieldbus Coupler]
//           modules: Module 1 (32 Byte Valve Unit (0x7F))
//         R10-VI12 (AES-D-BC-ECAT) [AES Fieldbus Coupler]
//           modules: Module 1 (32 Byte Valve Unit (0x7F))
//         R10_SAFETY (Flexi Soft EtherCAT Gateway) [Flexi Soft EtherCAT Gateway]
//       R10_A3 (EK1122) [EK1122 2 port EtherCAT junction]
//         R10-AB00 (EPP1322-0001) [EPP1322-0001 3 port EtherCAT P gateway]
//           R10-AB9 (EPP1008-0001) [EPP1008-0001 8 Ch. Dig. Input 24V, 3ms, M8]
//           R10-AB10 (EPP1008-0001) [EPP1008-0001 8 Ch. Dig. Input 24V, 3ms, M8]
//           R10-AB01 (EPP1332-0001) [EPP1332-0001 3 port EtherCAT P junction, power refreshing]
//             R10-ABT8 (EPP1008-0001) [EPP1008-0001 8 Ch. Dig. Input 24V, 3ms, M8]
//             R10-ABT9 (EPP1008-0001) [EPP1008-0001 8 Ch. Dig. Input 24V, 3ms, M8]
//             R10-ABT10 (EPP1008-0001) [EPP1008-0001 8 Ch. Dig. Input 24V, 3ms, M8]
//             R10-ABT11 (EPP1008-0001) [EPP1008-0001 8 Ch. Dig. Input 24V, 3ms, M8]
//             R10-ABT12 (EPP1008-0001) [EPP1008-0001 8 Ch. Dig. Input 24V, 3ms, M8]
//           R10-ABT7 (EPP1008-0001) [EPP1008-0001 8 Ch. Dig. Input 24V, 3ms, M8]
//           R10-ABT6 (EPP1008-0001) [EPP1008-0001 8 Ch. Dig. Input 24V, 3ms, M8]
//           R10-ABT5 (EPP1008-0001) [EPP1008-0001 8 Ch. Dig. Input 24V, 3ms, M8]
//           R10-ABT4 (EPP1008-0001) [EPP1008-0001 8 Ch. Dig. Input 24V, 3ms, M8]
//           R10-ABT3 (EPP1008-0001) [EPP1008-0001 8 Ch. Dig. Input 24V, 3ms, M8]
//           R10-ABT2 (EPP1008-0001) [EPP1008-0001 8 Ch. Dig. Input 24V, 3ms, M8]
//           R10-ABT1 (EPP1008-0001) [EPP1008-0001 8 Ch. Dig. Input 24V, 3ms, M8]
//         R10-AB1 (EPP1008-0001) [EPP1008-0001 8 Ch. Dig. Input 24V, 3ms, M8]
//         R10-AB2 (EPP1008-0001) [EPP1008-0001 8 Ch. Dig. Input 24V, 3ms, M8]
//         R10-AB3 (EPP1008-0001) [EPP1008-0001 8 Ch. Dig. Input 24V, 3ms, M8]
//         R10-AB4 (EPP1008-0001) [EPP1008-0001 8 Ch. Dig. Input 24V, 3ms, M8]
//         R10-AB5 (EPP1008-0001) [EPP1008-0001 8 Ch. Dig. Input 24V, 3ms, M8]
//         R10-AB6 (EPP1008-0001) [EPP1008-0001 8 Ch. Dig. Input 24V, 3ms, M8]
//         R10-AB02 (EPP1332-0001) [EPP1332-0001 3 port EtherCAT P junction, power refreshing]
//         R10-AB7 (EPP1008-0001) [EPP1008-0001 8 Ch. Dig. Input 24V, 3ms, M8]
//         R10-AB8 (EPP1008-0001) [EPP1008-0001 8 Ch. Dig. Input 24V, 3ms, M8]
//         R10-AB11 (EPP2308-0001) [EPP2308-0001 4 Ch. Dig. In, 3ms, 4 Ch. Dig. Out 24V, 0,5A, M8]
//         R10-AB12 (EPP2308-0001) [EPP2308-0001 4 Ch. Dig. In, 3ms, 4 Ch. Dig. Out 24V, 0,5A, M8]
//         R10-AB13 (EPP2308-0001) [EPP2308-0001 4 Ch. Dig. In, 3ms, 4 Ch. Dig. Out 24V, 0,5A, M8]
//       R10_A4 (EL6631) [EL6631 PROFINET IO Controller]
//       R10_A4 (EL7041-1000) [EL7041-1000 1Ch. Stepper motor output stage (50V, 5A, standard)]
//       R10_A5 (EL1809) [EL1809 16Ch. Dig. Input 24V, 3ms]
//       R10_A6 (EL2809) [EL2809 16Ch. Dig. Output 24V, 0.5A]
//       R10_A7 (EL2809) [EL2809 16Ch. Dig. Output 24V, 0.5A]
//       R10_A8 (EL3024) [EL3024 4Ch. Ana. Input 4-20mA DIFF]
//       R10_A9 (EL1809) [EL1809 16Ch. Dig. Input 24V, 3ms]
//       R10_A10 (EL2809) [EL2809 16Ch. Dig. Output 24V, 0.5A]
//       R10_EndTerminal (EL9011) [EL9011 End Terminal]
//   DEVICE Device 5 (EtherCAT) (disabled), AmsNetId 172.20.10.110.6.1
//     Term 279 (EK1100) [EK1100 EtherCAT Coupler (2A E-Bus)]
//       Term 280 (EL1809) [EL1809 16Ch. Dig. Input 24V, 3ms]
//       Term 281 (EL1809) [EL1809 16Ch. Dig. Input 24V, 3ms]
//       Term 282 (EL1809) [EL1809 16Ch. Dig. Input 24V, 3ms]
//       Term 283 (EL1809) [EL1809 16Ch. Dig. Input 24V, 3ms]
//       Term 284 (EL1809) [EL1809 16Ch. Dig. Input 24V, 3ms]
//       Term 312 (EL1809) [EL1809 16Ch. Dig. Input 24V, 3ms]
//       Term 320 (EL1809) [EL1809 16Ch. Dig. Input 24V, 3ms]
//       Term 321 (EL1809) [EL1809 16Ch. Dig. Input 24V, 3ms]
//       Term 322 (EL1809) [EL1809 16Ch. Dig. Input 24V, 3ms]
//       Term 323 (EL1809) [EL1809 16Ch. Dig. Input 24V, 3ms]
//       Term 324 (EL1809) [EL1809 16Ch. Dig. Input 24V, 3ms]
//       Term 325 (EL1809) [EL1809 16Ch. Dig. Input 24V, 3ms]
//       Term 326 (EL1809) [EL1809 16Ch. Dig. Input 24V, 3ms]
//       Term 327 (EL1809) [EL1809 16Ch. Dig. Input 24V, 3ms]
//       Term 328 (EL1809) [EL1809 16Ch. Dig. Input 24V, 3ms]
//       Term 329 (EL1809) [EL1809 16Ch. Dig. Input 24V, 3ms]
//       Term 331 (EL1809) [EL1809 16Ch. Dig. Input 24V, 3ms]
//       Term 332 (EL1809) [EL1809 16Ch. Dig. Input 24V, 3ms]
//       Term 333 (EL1809) [EL1809 16Ch. Dig. Input 24V, 3ms]
//       Term 334 (EL1809) [EL1809 16Ch. Dig. Input 24V, 3ms]
//       Term 335 (EL1809) [EL1809 16Ch. Dig. Input 24V, 3ms]
//       Term 336 (EL1809) [EL1809 16Ch. Dig. Input 24V, 3ms]
//       Term 337 (EL1809) [EL1809 16Ch. Dig. Input 24V, 3ms]
//       Term 338 (EL1809) [EL1809 16Ch. Dig. Input 24V, 3ms]
//       Term 339 (EL1809) [EL1809 16Ch. Dig. Input 24V, 3ms]
//       Term 340 (EL1809) [EL1809 16Ch. Dig. Input 24V, 3ms]
//       Term 341 (EL1809) [EL1809 16Ch. Dig. Input 24V, 3ms]
//       Term 342 (EL1809) [EL1809 16Ch. Dig. Input 24V, 3ms]
//       Term 343 (EL1809) [EL1809 16Ch. Dig. Input 24V, 3ms]
//       Term 344 (EL1809) [EL1809 16Ch. Dig. Input 24V, 3ms]
//       Term 345 (EL1809) [EL1809 16Ch. Dig. Input 24V, 3ms]
//       Term 346 (EL1809) [EL1809 16Ch. Dig. Input 24V, 3ms]
//       Term 347 (EL1809) [EL1809 16Ch. Dig. Input 24V, 3ms]
//       Term 348 (EL1809) [EL1809 16Ch. Dig. Input 24V, 3ms]
//       Term 360 (EL1809) [EL1809 16Ch. Dig. Input 24V, 3ms]
//       Term 361 (EL1809) [EL1809 16Ch. Dig. Input 24V, 3ms]
//       Term 362 (EL1809) [EL1809 16Ch. Dig. Input 24V, 3ms]
//       Term 363 (EL1809) [EL1809 16Ch. Dig. Input 24V, 3ms]
//       Term 364 (EL1809) [EL1809 16Ch. Dig. Input 24V, 3ms]
//       Term 365 (EL1809) [EL1809 16Ch. Dig. Input 24V, 3ms]
//       Term 366 (EL1809) [EL1809 16Ch. Dig. Input 24V, 3ms]
//       Term 367 (EL1809) [EL1809 16Ch. Dig. Input 24V, 3ms]
//       Term 368 (EL1809) [EL1809 16Ch. Dig. Input 24V, 3ms]
//       Term 370 (EL1809) [EL1809 16Ch. Dig. Input 24V, 3ms]
//       Term 371 (EL1809) [EL1809 16Ch. Dig. Input 24V, 3ms]
//       Term 372 (EL1809) [EL1809 16Ch. Dig. Input 24V, 3ms]
//       Term 373 (EL1809) [EL1809 16Ch. Dig. Input 24V, 3ms]
//       Term 374 (EL1809) [EL1809 16Ch. Dig. Input 24V, 3ms]
//       Term 375 (EL1809) [EL1809 16Ch. Dig. Input 24V, 3ms]
//       Term 376 (EL1809) [EL1809 16Ch. Dig. Input 24V, 3ms]
//       Term 377 (EL1809) [EL1809 16Ch. Dig. Input 24V, 3ms]
//       Term 378 (EL1809) [EL1809 16Ch. Dig. Input 24V, 3ms]
//       Term 380 (EL1809) [EL1809 16Ch. Dig. Input 24V, 3ms]
//       Term 381 (EL1809) [EL1809 16Ch. Dig. Input 24V, 3ms]
//       Term 382 (EL1809) [EL1809 16Ch. Dig. Input 24V, 3ms]
//       Term 383 (EL1809) [EL1809 16Ch. Dig. Input 24V, 3ms]
//       Term 384 (EL1809) [EL1809 16Ch. Dig. Input 24V, 3ms]
//       Term 385 (EL1809) [EL1809 16Ch. Dig. Input 24V, 3ms]
//       Term 386 (EL1809) [EL1809 16Ch. Dig. Input 24V, 3ms]
//       Term 387 (EL1809) [EL1809 16Ch. Dig. Input 24V, 3ms]
//       Term 388 (EL1809) [EL1809 16Ch. Dig. Input 24V, 3ms]
//       Term 389 (EL1809) [EL1809 16Ch. Dig. Input 24V, 3ms]
//       Term 390 (EL1809) [EL1809 16Ch. Dig. Input 24V, 3ms]
//       Term 391 (EL1809) [EL1809 16Ch. Dig. Input 24V, 3ms]
//       Term 392 (EL1809) [EL1809 16Ch. Dig. Input 24V, 3ms]
//       Term 393 (EL1809) [EL1809 16Ch. Dig. Input 24V, 3ms]
//       Term 394 (EL1809) [EL1809 16Ch. Dig. Input 24V, 3ms]
//       Term 395 (EL1809) [EL1809 16Ch. Dig. Input 24V, 3ms]
//       Term 396 (EL1809) [EL1809 16Ch. Dig. Input 24V, 3ms]
//       Term 397 (EL1809) [EL1809 16Ch. Dig. Input 24V, 3ms]
//       Term 398 (EL1809) [EL1809 16Ch. Dig. Input 24V, 3ms]
//       Term 399 (EL1809) [EL1809 16Ch. Dig. Input 24V, 3ms]
//       Term 400 (EL1809) [EL1809 16Ch. Dig. Input 24V, 3ms]
//       Term 401 (EL1809) [EL1809 16Ch. Dig. Input 24V, 3ms]
//       Term 402 (EL1809) [EL1809 16Ch. Dig. Input 24V, 3ms]
//       Term 403 (EL1809) [EL1809 16Ch. Dig. Input 24V, 3ms]
//       Term 404 (EL1809) [EL1809 16Ch. Dig. Input 24V, 3ms]
//       Term 405 (EL1809) [EL1809 16Ch. Dig. Input 24V, 3ms]
//       Term 406 (EL1809) [EL1809 16Ch. Dig. Input 24V, 3ms]
//       Term 407 (EL1809) [EL1809 16Ch. Dig. Input 24V, 3ms]
//       Term 408 (EL1809) [EL1809 16Ch. Dig. Input 24V, 3ms]
//       Term 409 (EL1809) [EL1809 16Ch. Dig. Input 24V, 3ms]
//       Term 410 (EL1809) [EL1809 16Ch. Dig. Input 24V, 3ms]
//       Term 414 (EL1809) [EL1809 16Ch. Dig. Input 24V, 3ms]
//       Term 415 (EL1809) [EL1809 16Ch. Dig. Input 24V, 3ms]
//       Term 416 (EL1809) [EL1809 16Ch. Dig. Input 24V, 3ms]
//       Term 417 (EL1809) [EL1809 16Ch. Dig. Input 24V, 3ms]
//       Term 418 (EL1809) [EL1809 16Ch. Dig. Input 24V, 3ms]
//       Term 419 (EL1809) [EL1809 16Ch. Dig. Input 24V, 3ms]
//       Term 420 (EL1809) [EL1809 16Ch. Dig. Input 24V, 3ms]
//       Term 421 (EL1809) [EL1809 16Ch. Dig. Input 24V, 3ms]
//       Term 422 (EL1809) [EL1809 16Ch. Dig. Input 24V, 3ms]
//       Term 423 (EL1809) [EL1809 16Ch. Dig. Input 24V, 3ms]
//       Term 424 (EL1809) [EL1809 16Ch. Dig. Input 24V, 3ms]
//       Term 425 (EL1809) [EL1809 16Ch. Dig. Input 24V, 3ms]
//       Term 426 (EL1809) [EL1809 16Ch. Dig. Input 24V, 3ms]
//       Term 427 (EL1809) [EL1809 16Ch. Dig. Input 24V, 3ms]
//       Term 428 (EL1809) [EL1809 16Ch. Dig. Input 24V, 3ms]
//       Term 429 (EL1809) [EL1809 16Ch. Dig. Input 24V, 3ms]
//       Term 448 (EL1809) [EL1809 16Ch. Dig. Input 24V, 3ms]
//       Term 495 (EK1110) [EK1110 EtherCAT extension]
//     Term 554 (EK1100) [EK1100 EtherCAT Coupler (2A E-Bus)]
//       Term 645 (EL1809) [EL1809 16Ch. Dig. Input 24V, 3ms]
//       Term 646 (EL1809) [EL1809 16Ch. Dig. Input 24V, 3ms]
//       Term 647 (EL1809) [EL1809 16Ch. Dig. Input 24V, 3ms]
//       Term 648 (EL1809) [EL1809 16Ch. Dig. Input 24V, 3ms]
//       Term 649 (EL1809) [EL1809 16Ch. Dig. Input 24V, 3ms]
//       Term 650 (EL1809) [EL1809 16Ch. Dig. Input 24V, 3ms]
//       Term 651 (EL1809) [EL1809 16Ch. Dig. Input 24V, 3ms]
//       Term 652 (EL1809) [EL1809 16Ch. Dig. Input 24V, 3ms]
//       Term 653 (EL1809) [EL1809 16Ch. Dig. Input 24V, 3ms]
//       Term 654 (EL1809) [EL1809 16Ch. Dig. Input 24V, 3ms]
//       Term 655 (EL1809) [EL1809 16Ch. Dig. Input 24V, 3ms]
//       Term 656 (EL1809) [EL1809 16Ch. Dig. Input 24V, 3ms]
//       Term 657 (EL1809) [EL1809 16Ch. Dig. Input 24V, 3ms]
//       Term 658 (EL1809) [EL1809 16Ch. Dig. Input 24V, 3ms]
//       Term 659 (EL1809) [EL1809 16Ch. Dig. Input 24V, 3ms]
//       Term 660 (EL1809) [EL1809 16Ch. Dig. Input 24V, 3ms]
//       Term 661 (EL1809) [EL1809 16Ch. Dig. Input 24V, 3ms]
//       Term 662 (EL1809) [EL1809 16Ch. Dig. Input 24V, 3ms]
//       Term 663 (EL1809) [EL1809 16Ch. Dig. Input 24V, 3ms]
//       Term 664 (EL1809) [EL1809 16Ch. Dig. Input 24V, 3ms]
//       Term 665 (EL1809) [EL1809 16Ch. Dig. Input 24V, 3ms]
//       Term 666 (EL1809) [EL1809 16Ch. Dig. Input 24V, 3ms]
//       Term 667 (EL1809) [EL1809 16Ch. Dig. Input 24V, 3ms]
//       Term 668 (EL1809) [EL1809 16Ch. Dig. Input 24V, 3ms]
//       Term 669 (EL1809) [EL1809 16Ch. Dig. Input 24V, 3ms]
//       Term 670 (EL1809) [EL1809 16Ch. Dig. Input 24V, 3ms]
//       Term 671 (EL1809) [EL1809 16Ch. Dig. Input 24V, 3ms]
//       Term 672 (EL1809) [EL1809 16Ch. Dig. Input 24V, 3ms]
//       Term 673 (EL1809) [EL1809 16Ch. Dig. Input 24V, 3ms]
//       Term 674 (EL1809) [EL1809 16Ch. Dig. Input 24V, 3ms]
//       Term 676 (EL1809) [EL1809 16Ch. Dig. Input 24V, 3ms]
//       Term 677 (EL1809) [EL1809 16Ch. Dig. Input 24V, 3ms]
//       Term 678 (EL1809) [EL1809 16Ch. Dig. Input 24V, 3ms]
//       Term 679 (EL1809) [EL1809 16Ch. Dig. Input 24V, 3ms]
//       Term 680 (EL1809) [EL1809 16Ch. Dig. Input 24V, 3ms]
//       Term 681 (EL1809) [EL1809 16Ch. Dig. Input 24V, 3ms]
//       Term 682 (EL1809) [EL1809 16Ch. Dig. Input 24V, 3ms]
//       Term 683 (EL1809) [EL1809 16Ch. Dig. Input 24V, 3ms]
//       Term 684 (EL1809) [EL1809 16Ch. Dig. Input 24V, 3ms]
//       Term 685 (EL1809) [EL1809 16Ch. Dig. Input 24V, 3ms]
//       Term 686 (EL1809) [EL1809 16Ch. Dig. Input 24V, 3ms]
//       Term 687 (EL1809) [EL1809 16Ch. Dig. Input 24V, 3ms]
//       Term 688 (EL1809) [EL1809 16Ch. Dig. Input 24V, 3ms]
//       Term 689 (EL1809) [EL1809 16Ch. Dig. Input 24V, 3ms]
//       Term 690 (EL1809) [EL1809 16Ch. Dig. Input 24V, 3ms]
//       Term 691 (EL1809) [EL1809 16Ch. Dig. Input 24V, 3ms]
//       Term 692 (EL1809) [EL1809 16Ch. Dig. Input 24V, 3ms]
//       Term 693 (EL1809) [EL1809 16Ch. Dig. Input 24V, 3ms]
//       Term 694 (EL1809) [EL1809 16Ch. Dig. Input 24V, 3ms]
//       Term 695 (EL1809) [EL1809 16Ch. Dig. Input 24V, 3ms]
//       Term 696 (EL1809) [EL1809 16Ch. Dig. Input 24V, 3ms]
//       Term 697 (EL1809) [EL1809 16Ch. Dig. Input 24V, 3ms]
//       Term 698 (EL1809) [EL1809 16Ch. Dig. Input 24V, 3ms]
//       Term 699 (EL1809) [EL1809 16Ch. Dig. Input 24V, 3ms]
//       Term 700 (EL1809) [EL1809 16Ch. Dig. Input 24V, 3ms]
//       Term 701 (EL1809) [EL1809 16Ch. Dig. Input 24V, 3ms]
//       Term 702 (EL1809) [EL1809 16Ch. Dig. Input 24V, 3ms]
//       Term 703 (EL1809) [EL1809 16Ch. Dig. Input 24V, 3ms]
//       Term 704 (EL1809) [EL1809 16Ch. Dig. Input 24V, 3ms]
//       Term 705 (EL1809) [EL1809 16Ch. Dig. Input 24V, 3ms]
//       Term 706 (EL1809) [EL1809 16Ch. Dig. Input 24V, 3ms]
//       Term 707 (EL1809) [EL1809 16Ch. Dig. Input 24V, 3ms]
//       Term 709 (EL1809) [EL1809 16Ch. Dig. Input 24V, 3ms]
//       Term 710 (EL1809) [EL1809 16Ch. Dig. Input 24V, 3ms]
//       Term 711 (EL1809) [EL1809 16Ch. Dig. Input 24V, 3ms]
//       Term 712 (EL1809) [EL1809 16Ch. Dig. Input 24V, 3ms]
//       Term 713 (EL1809) [EL1809 16Ch. Dig. Input 24V, 3ms]
//       Term 714 (EL1809) [EL1809 16Ch. Dig. Input 24V, 3ms]
//       Term 715 (EL1809) [EL1809 16Ch. Dig. Input 24V, 3ms]
//       Term 716 (EL1809) [EL1809 16Ch. Dig. Input 24V, 3ms]
//       Term 717 (EL1809) [EL1809 16Ch. Dig. Input 24V, 3ms]
//       Term 718 (EL1809) [EL1809 16Ch. Dig. Input 24V, 3ms]
//       Term 719 (EL1809) [EL1809 16Ch. Dig. Input 24V, 3ms]
//       Term 720 (EL1809) [EL1809 16Ch. Dig. Input 24V, 3ms]
//       Term 721 (EL1809) [EL1809 16Ch. Dig. Input 24V, 3ms]
//       Term 722 (EL1809) [EL1809 16Ch. Dig. Input 24V, 3ms]
//       Term 723 (EL1809) [EL1809 16Ch. Dig. Input 24V, 3ms]
//       Term 724 (EL1809) [EL1809 16Ch. Dig. Input 24V, 3ms]
//       Term 725 (EL1809) [EL1809 16Ch. Dig. Input 24V, 3ms]
//       Term 726 (EL1809) [EL1809 16Ch. Dig. Input 24V, 3ms]
//       Term 727 (EL1809) [EL1809 16Ch. Dig. Input 24V, 3ms]
//       Term 728 (EL1809) [EL1809 16Ch. Dig. Input 24V, 3ms]
//       Term 729 (EL1809) [EL1809 16Ch. Dig. Input 24V, 3ms]
//       Term 730 (EL1809) [EL1809 16Ch. Dig. Input 24V, 3ms]
//       Term 731 (EL1809) [EL1809 16Ch. Dig. Input 24V, 3ms]
//       Term 732 (EL1809) [EL1809 16Ch. Dig. Input 24V, 3ms]
//       Term 733 (EL1809) [EL1809 16Ch. Dig. Input 24V, 3ms]
//       Term 734 (EL1809) [EL1809 16Ch. Dig. Input 24V, 3ms]
//       Term 735 (EL1809) [EL1809 16Ch. Dig. Input 24V, 3ms]
//       Term 736 (EL1809) [EL1809 16Ch. Dig. Input 24V, 3ms]
//       Term 737 (EL1809) [EL1809 16Ch. Dig. Input 24V, 3ms]
//       Term 738 (EL1809) [EL1809 16Ch. Dig. Input 24V, 3ms]
//       Term 739 (EL1809) [EL1809 16Ch. Dig. Input 24V, 3ms]
//       Term 740 (EL1809) [EL1809 16Ch. Dig. Input 24V, 3ms]
//       Term 741 (EL1809) [EL1809 16Ch. Dig. Input 24V, 3ms]
//       Term 742 (EL1809) [EL1809 16Ch. Dig. Input 24V, 3ms]
//       Term 743 (EL1809) [EL1809 16Ch. Dig. Input 24V, 3ms]
//       Term 744 (EL1809) [EL1809 16Ch. Dig. Input 24V, 3ms]
//       Term 745 (EL1809) [EL1809 16Ch. Dig. Input 24V, 3ms]
//       Term 746 (EL1809) [EL1809 16Ch. Dig. Input 24V, 3ms]
//       Term 747 (EK1110) [EK1110 EtherCAT extension]
//     Term 748 (EK1100) [EK1100 EtherCAT Coupler (2A E-Bus)]
//       Term 749 (EL1809) [EL1809 16Ch. Dig. Input 24V, 3ms]
//       Term 750 (EL1809) [EL1809 16Ch. Dig. Input 24V, 3ms]
//       Term 751 (EL1809) [EL1809 16Ch. Dig. Input 24V, 3ms]
//       Term 752 (EL1809) [EL1809 16Ch. Dig. Input 24V, 3ms]
//       Term 753 (EL1809) [EL1809 16Ch. Dig. Input 24V, 3ms]
//       Term 754 (EL1809) [EL1809 16Ch. Dig. Input 24V, 3ms]
//       Term 755 (EL1809) [EL1809 16Ch. Dig. Input 24V, 3ms]
//       Term 756 (EL1809) [EL1809 16Ch. Dig. Input 24V, 3ms]
//       Term 757 (EL1809) [EL1809 16Ch. Dig. Input 24V, 3ms]
//       Term 758 (EL1809) [EL1809 16Ch. Dig. Input 24V, 3ms]
//       Term 759 (EL1809) [EL1809 16Ch. Dig. Input 24V, 3ms]
//       Term 760 (EL1809) [EL1809 16Ch. Dig. Input 24V, 3ms]
//       Term 761 (EL1809) [EL1809 16Ch. Dig. Input 24V, 3ms]
//       Term 762 (EL1809) [EL1809 16Ch. Dig. Input 24V, 3ms]
//       Term 763 (EL1809) [EL1809 16Ch. Dig. Input 24V, 3ms]
//       Term 764 (EL1809) [EL1809 16Ch. Dig. Input 24V, 3ms]
//       Term 765 (EL1809) [EL1809 16Ch. Dig. Input 24V, 3ms]
//       Term 766 (EL1809) [EL1809 16Ch. Dig. Input 24V, 3ms]
//       Term 767 (EL1809) [EL1809 16Ch. Dig. Input 24V, 3ms]
//       Term 768 (EL1809) [EL1809 16Ch. Dig. Input 24V, 3ms]
//       Term 769 (EL1809) [EL1809 16Ch. Dig. Input 24V, 3ms]
//       Term 770 (EL1809) [EL1809 16Ch. Dig. Input 24V, 3ms]
//       Term 771 (EL1809) [EL1809 16Ch. Dig. Input 24V, 3ms]
//       Term 772 (EL1809) [EL1809 16Ch. Dig. Input 24V, 3ms]
//       Term 773 (EL1809) [EL1809 16Ch. Dig. Input 24V, 3ms]
//       Term 774 (EL1809) [EL1809 16Ch. Dig. Input 24V, 3ms]
//       Term 775 (EL1809) [EL1809 16Ch. Dig. Input 24V, 3ms]
//       Term 776 (EL1809) [EL1809 16Ch. Dig. Input 24V, 3ms]
//       Term 777 (EL1809) [EL1809 16Ch. Dig. Input 24V, 3ms]
//       Term 778 (EL1809) [EL1809 16Ch. Dig. Input 24V, 3ms]
//       Term 779 (EL1809) [EL1809 16Ch. Dig. Input 24V, 3ms]
//       Term 780 (EL1809) [EL1809 16Ch. Dig. Input 24V, 3ms]
//       Term 781 (EL1809) [EL1809 16Ch. Dig. Input 24V, 3ms]
//       Term 782 (EL1809) [EL1809 16Ch. Dig. Input 24V, 3ms]
//       Term 783 (EL1809) [EL1809 16Ch. Dig. Input 24V, 3ms]
//       Term 784 (EL1809) [EL1809 16Ch. Dig. Input 24V, 3ms]
//       Term 785 (EL1809) [EL1809 16Ch. Dig. Input 24V, 3ms]
//       Term 786 (EL1809) [EL1809 16Ch. Dig. Input 24V, 3ms]
//       Term 787 (EL1809) [EL1809 16Ch. Dig. Input 24V, 3ms]
//       Term 788 (EL1809) [EL1809 16Ch. Dig. Input 24V, 3ms]
//       Term 789 (EL1809) [EL1809 16Ch. Dig. Input 24V, 3ms]
//       Term 790 (EL1809) [EL1809 16Ch. Dig. Input 24V, 3ms]
//       Term 791 (EL1809) [EL1809 16Ch. Dig. Input 24V, 3ms]
//       Term 792 (EL1809) [EL1809 16Ch. Dig. Input 24V, 3ms]
//       Term 793 (EL1809) [EL1809 16Ch. Dig. Input 24V, 3ms]
//       Term 794 (EL1809) [EL1809 16Ch. Dig. Input 24V, 3ms]
//       Term 795 (EL1809) [EL1809 16Ch. Dig. Input 24V, 3ms]
//       Term 796 (EL1809) [EL1809 16Ch. Dig. Input 24V, 3ms]
//       Term 798 (EL1809) [EL1809 16Ch. Dig. Input 24V, 3ms]
//       Term 799 (EL1809) [EL1809 16Ch. Dig. Input 24V, 3ms]
//       Term 800 (EL1809) [EL1809 16Ch. Dig. Input 24V, 3ms]
//       Term 801 (EL1809) [EL1809 16Ch. Dig. Input 24V, 3ms]
//       Term 802 (EL1809) [EL1809 16Ch. Dig. Input 24V, 3ms]
//       Term 803 (EL1809) [EL1809 16Ch. Dig. Input 24V, 3ms]
//       Term 804 (EL1809) [EL1809 16Ch. Dig. Input 24V, 3ms]
//       Term 805 (EL1809) [EL1809 16Ch. Dig. Input 24V, 3ms]
//       Term 806 (EL1809) [EL1809 16Ch. Dig. Input 24V, 3ms]
//       Term 807 (EL1809) [EL1809 16Ch. Dig. Input 24V, 3ms]
//       Term 808 (EL1809) [EL1809 16Ch. Dig. Input 24V, 3ms]
//       Term 809 (EL1809) [EL1809 16Ch. Dig. Input 24V, 3ms]
//       Term 810 (EL1809) [EL1809 16Ch. Dig. Input 24V, 3ms]
//       Term 811 (EL1809) [EL1809 16Ch. Dig. Input 24V, 3ms]
//       Term 812 (EL1809) [EL1809 16Ch. Dig. Input 24V, 3ms]
//       Term 813 (EL1809) [EL1809 16Ch. Dig. Input 24V, 3ms]
//       Term 814 (EL1809) [EL1809 16Ch. Dig. Input 24V, 3ms]
//       Term 815 (EL1809) [EL1809 16Ch. Dig. Input 24V, 3ms]
//       Term 816 (EL1809) [EL1809 16Ch. Dig. Input 24V, 3ms]
//       Term 817 (EL1809) [EL1809 16Ch. Dig. Input 24V, 3ms]
//       Term 818 (EL1809) [EL1809 16Ch. Dig. Input 24V, 3ms]
//       Term 819 (EL1809) [EL1809 16Ch. Dig. Input 24V, 3ms]
//       Term 820 (EL1809) [EL1809 16Ch. Dig. Input 24V, 3ms]
//       Term 821 (EL1809) [EL1809 16Ch. Dig. Input 24V, 3ms]
//       Term 822 (EL1809) [EL1809 16Ch. Dig. Input 24V, 3ms]
//       Term 823 (EL1809) [EL1809 16Ch. Dig. Input 24V, 3ms]
//       Term 824 (EL1809) [EL1809 16Ch. Dig. Input 24V, 3ms]
//       Term 825 (EL1809) [EL1809 16Ch. Dig. Input 24V, 3ms]
//       Term 826 (EL1809) [EL1809 16Ch. Dig. Input 24V, 3ms]
//       Term 827 (EL1809) [EL1809 16Ch. Dig. Input 24V, 3ms]
//       Term 828 (EL1809) [EL1809 16Ch. Dig. Input 24V, 3ms]
//       Term 859 (EL1809) [EL1809 16Ch. Dig. Input 24V, 3ms]
//       Term 860 (EL1809) [EL1809 16Ch. Dig. Input 24V, 3ms]
//       Term 861 (EL1809) [EL1809 16Ch. Dig. Input 24V, 3ms]
//       Term 862 (EL1809) [EL1809 16Ch. Dig. Input 24V, 3ms]
//       Term 863 (EL1809) [EL1809 16Ch. Dig. Input 24V, 3ms]
//       Term 864 (EL1809) [EL1809 16Ch. Dig. Input 24V, 3ms]
//       Term 865 (EL1809) [EL1809 16Ch. Dig. Input 24V, 3ms]
//       Term 866 (EL1809) [EL1809 16Ch. Dig. Input 24V, 3ms]
//       Term 867 (EL1809) [EL1809 16Ch. Dig. Input 24V, 3ms]
//       Term 868 (EL1809) [EL1809 16Ch. Dig. Input 24V, 3ms]
//       Term 869 (EL1809) [EL1809 16Ch. Dig. Input 24V, 3ms]
//       Term 870 (EL1809) [EL1809 16Ch. Dig. Input 24V, 3ms]
//       Term 871 (EL1809) [EL1809 16Ch. Dig. Input 24V, 3ms]
//       Term 872 (EL1809) [EL1809 16Ch. Dig. Input 24V, 3ms]
//       Term 873 (EL1809) [EL1809 16Ch. Dig. Input 24V, 3ms]
//       Term 874 (EL1809) [EL1809 16Ch. Dig. Input 24V, 3ms]
//       Term 875 (EL1809) [EL1809 16Ch. Dig. Input 24V, 3ms]
//       Term 876 (EL1809) [EL1809 16Ch. Dig. Input 24V, 3ms]
//       Term 877 (EL1809) [EL1809 16Ch. Dig. Input 24V, 3ms]
//       Term 878 (EL1809) [EL1809 16Ch. Dig. Input 24V, 3ms]
//       Term 879 (EL1809) [EL1809 16Ch. Dig. Input 24V, 3ms]
//       Term 880 (EK1110) [EK1110 EtherCAT extension]
//     Term 881 (EK1100) [EK1100 EtherCAT Coupler (2A E-Bus)]
//       Term 882 (EL1809) [EL1809 16Ch. Dig. Input 24V, 3ms]
//       Term 883 (EL1809) [EL1809 16Ch. Dig. Input 24V, 3ms]
//       Term 884 (EL1809) [EL1809 16Ch. Dig. Input 24V, 3ms]
//       Term 885 (EL1809) [EL1809 16Ch. Dig. Input 24V, 3ms]
//       Term 886 (EL1809) [EL1809 16Ch. Dig. Input 24V, 3ms]
//       Term 887 (EL1809) [EL1809 16Ch. Dig. Input 24V, 3ms]
//       Term 888 (EL1809) [EL1809 16Ch. Dig. Input 24V, 3ms]
//       Term 889 (EL1809) [EL1809 16Ch. Dig. Input 24V, 3ms]
//       Term 890 (EL1809) [EL1809 16Ch. Dig. Input 24V, 3ms]
//       Term 891 (EL1809) [EL1809 16Ch. Dig. Input 24V, 3ms]
//       Term 892 (EL1809) [EL1809 16Ch. Dig. Input 24V, 3ms]
//       Term 893 (EL1809) [EL1809 16Ch. Dig. Input 24V, 3ms]
//       Term 894 (EL1809) [EL1809 16Ch. Dig. Input 24V, 3ms]
//       Term 895 (EL1809) [EL1809 16Ch. Dig. Input 24V, 3ms]
//       Term 896 (EL1809) [EL1809 16Ch. Dig. Input 24V, 3ms]
//       Term 897 (EL1809) [EL1809 16Ch. Dig. Input 24V, 3ms]
//       Term 898 (EL1809) [EL1809 16Ch. Dig. Input 24V, 3ms]
//       Term 899 (EL1809) [EL1809 16Ch. Dig. Input 24V, 3ms]
//       Term 900 (EL1809) [EL1809 16Ch. Dig. Input 24V, 3ms]
//       Term 901 (EL1809) [EL1809 16Ch. Dig. Input 24V, 3ms]
//       Term 902 (EL1809) [EL1809 16Ch. Dig. Input 24V, 3ms]
//       Term 903 (EL1809) [EL1809 16Ch. Dig. Input 24V, 3ms]
//       Term 904 (EL1809) [EL1809 16Ch. Dig. Input 24V, 3ms]
//       Term 905 (EL1809) [EL1809 16Ch. Dig. Input 24V, 3ms]
//       Term 906 (EL1809) [EL1809 16Ch. Dig. Input 24V, 3ms]
//       Term 933 (EL1809) [EL1809 16Ch. Dig. Input 24V, 3ms]
//       Term 934 (EL1809) [EL1809 16Ch. Dig. Input 24V, 3ms]
//       Term 935 (EL1809) [EL1809 16Ch. Dig. Input 24V, 3ms]
//       Term 936 (EL1809) [EL1809 16Ch. Dig. Input 24V, 3ms]
//       Term 937 (EL1809) [EL1809 16Ch. Dig. Input 24V, 3ms]
//       Term 938 (EL1809) [EL1809 16Ch. Dig. Input 24V, 3ms]
//       Term 939 (EL1809) [EL1809 16Ch. Dig. Input 24V, 3ms]
//       Term 940 (EL1809) [EL1809 16Ch. Dig. Input 24V, 3ms]
//       Term 941 (EL1809) [EL1809 16Ch. Dig. Input 24V, 3ms]
//       Term 942 (EL1809) [EL1809 16Ch. Dig. Input 24V, 3ms]
//       Term 943 (EL1809) [EL1809 16Ch. Dig. Input 24V, 3ms]
//       Term 944 (EL1809) [EL1809 16Ch. Dig. Input 24V, 3ms]
//       Term 945 (EL1809) [EL1809 16Ch. Dig. Input 24V, 3ms]
//       Term 946 (EL1809) [EL1809 16Ch. Dig. Input 24V, 3ms]
//       Term 947 (EL1809) [EL1809 16Ch. Dig. Input 24V, 3ms]
//       Term 948 (EL1809) [EL1809 16Ch. Dig. Input 24V, 3ms]
//       Term 949 (EL1809) [EL1809 16Ch. Dig. Input 24V, 3ms]
//       Term 950 (EL1809) [EL1809 16Ch. Dig. Input 24V, 3ms]
//       Term 951 (EL1809) [EL1809 16Ch. Dig. Input 24V, 3ms]
//       Term 952 (EL1809) [EL1809 16Ch. Dig. Input 24V, 3ms]
//       Term 953 (EL1809) [EL1809 16Ch. Dig. Input 24V, 3ms]
//       Term 954 (EL1809) [EL1809 16Ch. Dig. Input 24V, 3ms]
//       Term 955 (EL1809) [EL1809 16Ch. Dig. Input 24V, 3ms]
//       Term 956 (EL1809) [EL1809 16Ch. Dig. Input 24V, 3ms]
//       Term 957 (EL1809) [EL1809 16Ch. Dig. Input 24V, 3ms]
//       Term 958 (EL1809) [EL1809 16Ch. Dig. Input 24V, 3ms]
//       Term 959 (EL1809) [EL1809 16Ch. Dig. Input 24V, 3ms]
//       Term 960 (EL1809) [EL1809 16Ch. Dig. Input 24V, 3ms]
//       Term 961 (EL1809) [EL1809 16Ch. Dig. Input 24V, 3ms]
//       Term 962 (EL1809) [EL1809 16Ch. Dig. Input 24V, 3ms]
//       Term 963 (EL1809) [EL1809 16Ch. Dig. Input 24V, 3ms]
//       Term 964 (EL1809) [EL1809 16Ch. Dig. Input 24V, 3ms]
//       Term 965 (EL1809) [EL1809 16Ch. Dig. Input 24V, 3ms]
//       Term 967 (EL1809) [EL1809 16Ch. Dig. Input 24V, 3ms]
//       Term 968 (EL1809) [EL1809 16Ch. Dig. Input 24V, 3ms]
//       Term 969 (EL1809) [EL1809 16Ch. Dig. Input 24V, 3ms]
//       Term 970 (EL1809) [EL1809 16Ch. Dig. Input 24V, 3ms]
//       Term 971 (EL1809) [EL1809 16Ch. Dig. Input 24V, 3ms]
//       Term 972 (EL1809) [EL1809 16Ch. Dig. Input 24V, 3ms]
//       Term 973 (EL1809) [EL1809 16Ch. Dig. Input 24V, 3ms]
//       Term 974 (EL1809) [EL1809 16Ch. Dig. Input 24V, 3ms]
//       Term 975 (EL1809) [EL1809 16Ch. Dig. Input 24V, 3ms]
//       Term 976 (EL1809) [EL1809 16Ch. Dig. Input 24V, 3ms]
//       Term 977 (EL1809) [EL1809 16Ch. Dig. Input 24V, 3ms]
//       Term 978 (EL1809) [EL1809 16Ch. Dig. Input 24V, 3ms]
//       Term 979 (EL1809) [EL1809 16Ch. Dig. Input 24V, 3ms]
//       Term 980 (EL1809) [EL1809 16Ch. Dig. Input 24V, 3ms]
//       Term 981 (EL1809) [EL1809 16Ch. Dig. Input 24V, 3ms]
//       Term 982 (EL1809) [EL1809 16Ch. Dig. Input 24V, 3ms]
//       Term 983 (EL1809) [EL1809 16Ch. Dig. Input 24V, 3ms]
//       Term 984 (EL1809) [EL1809 16Ch. Dig. Input 24V, 3ms]
//       Term 986 (EL1809) [EL1809 16Ch. Dig. Input 24V, 3ms]
//       Term 987 (EL1809) [EL1809 16Ch. Dig. Input 24V, 3ms]
//       Term 988 (EL1809) [EL1809 16Ch. Dig. Input 24V, 3ms]
//       Term 989 (EL1809) [EL1809 16Ch. Dig. Input 24V, 3ms]
//       Term 1025 (EL1809) [EL1809 16Ch. Dig. Input 24V, 3ms]
//       Term 1026 (EL1809) [EL1809 16Ch. Dig. Input 24V, 3ms]
//       Term 1027 (EL1809) [EL1809 16Ch. Dig. Input 24V, 3ms]
//       Term 1028 (EL1809) [EL1809 16Ch. Dig. Input 24V, 3ms]
//       Term 1029 (EL1809) [EL1809 16Ch. Dig. Input 24V, 3ms]
//       Term 1030 (EL1809) [EL1809 16Ch. Dig. Input 24V, 3ms]
//       Term 1031 (EL1809) [EL1809 16Ch. Dig. Input 24V, 3ms]
//       Term 1032 (EL1809) [EL1809 16Ch. Dig. Input 24V, 3ms]
//       Term 1033 (EL1809) [EL1809 16Ch. Dig. Input 24V, 3ms]
//       Term 1034 (EL1809) [EL1809 16Ch. Dig. Input 24V, 3ms]
//       Term 1035 (EL1809) [EL1809 16Ch. Dig. Input 24V, 3ms]
//       Term 1036 (EL1809) [EL1809 16Ch. Dig. Input 24V, 3ms]
//       Term 1038 (EL1809) [EL1809 16Ch. Dig. Input 24V, 3ms]
//       Term 1039 (EL1809) [EL1809 16Ch. Dig. Input 24V, 3ms]
//       Term 1040 (EL1809) [EL1809 16Ch. Dig. Input 24V, 3ms]
//       Term 1041 (EL1809) [EL1809 16Ch. Dig. Input 24V, 3ms]
//       Term 1042 (EL1809) [EL1809 16Ch. Dig. Input 24V, 3ms]
//       Term 1043 (EL1809) [EL1809 16Ch. Dig. Input 24V, 3ms]
//       Term 1044 (EL1809) [EL1809 16Ch. Dig. Input 24V, 3ms]
//       Term 1045 (EL1809) [EL1809 16Ch. Dig. Input 24V, 3ms]
//       Term 1046 (EK1110) [EK1110 EtherCAT extension]
//     Term 1047 (EK1100) [EK1100 EtherCAT Coupler (2A E-Bus)]
//       Term 1048 (EL1809) [EL1809 16Ch. Dig. Input 24V, 3ms]
//       Term 1049 (EL1809) [EL1809 16Ch. Dig. Input 24V, 3ms]
//       Term 1050 (EL1809) [EL1809 16Ch. Dig. Input 24V, 3ms]
//       Term 1051 (EL1809) [EL1809 16Ch. Dig. Input 24V, 3ms]
//       Term 1052 (EL1809) [EL1809 16Ch. Dig. Input 24V, 3ms]
//       Term 1053 (EL1809) [EL1809 16Ch. Dig. Input 24V, 3ms]
//       Term 1054 (EL1809) [EL1809 16Ch. Dig. Input 24V, 3ms]
//       Term 1055 (EL1809) [EL1809 16Ch. Dig. Input 24V, 3ms]
//       Term 1056 (EL1809) [EL1809 16Ch. Dig. Input 24V, 3ms]
//       Term 1057 (EL1809) [EL1809 16Ch. Dig. Input 24V, 3ms]
//       Term 1058 (EL1809) [EL1809 16Ch. Dig. Input 24V, 3ms]
//       Term 1059 (EL1809) [EL1809 16Ch. Dig. Input 24V, 3ms]
//       Term 1060 (EL1809) [EL1809 16Ch. Dig. Input 24V, 3ms]
//       Term 1061 (EL1809) [EL1809 16Ch. Dig. Input 24V, 3ms]
//       Term 1062 (EL1809) [EL1809 16Ch. Dig. Input 24V, 3ms]
//       Term 1063 (EL1809) [EL1809 16Ch. Dig. Input 24V, 3ms]
//       Term 1064 (EL1809) [EL1809 16Ch. Dig. Input 24V, 3ms]
//       Term 1065 (EL1809) [EL1809 16Ch. Dig. Input 24V, 3ms]
//       Term 1066 (EL1809) [EL1809 16Ch. Dig. Input 24V, 3ms]
//       Term 1068 (EL1809) [EL1809 16Ch. Dig. Input 24V, 3ms]
//       Term 1069 (EL1809) [EL1809 16Ch. Dig. Input 24V, 3ms]
//       Term 1070 (EL1809) [EL1809 16Ch. Dig. Input 24V, 3ms]
//       Term 1072 (EL1809) [EL1809 16Ch. Dig. Input 24V, 3ms]
//       Term 1073 (EL1809) [EL1809 16Ch. Dig. Input 24V, 3ms]
//       Term 1076 (EL1809) [EL1809 16Ch. Dig. Input 24V, 3ms]
//       Term 1077 (EL1809) [EL1809 16Ch. Dig. Input 24V, 3ms]
//       Term 1078 (EL1809) [EL1809 16Ch. Dig. Input 24V, 3ms]
//       Term 1081 (EL1809) [EL1809 16Ch. Dig. Input 24V, 3ms]
//       Term 1082 (EL1809) [EL1809 16Ch. Dig. Input 24V, 3ms]
//       Term 1083 (EL1809) [EL1809 16Ch. Dig. Input 24V, 3ms]
//       Term 1084 (EL1809) [EL1809 16Ch. Dig. Input 24V, 3ms]
//       Term 1085 (EL1809) [EL1809 16Ch. Dig. Input 24V, 3ms]
//       Term 1086 (EL1809) [EL1809 16Ch. Dig. Input 24V, 3ms]
//       Term 1087 (EL1809) [EL1809 16Ch. Dig. Input 24V, 3ms]
//       Term 1088 (EL1809) [EL1809 16Ch. Dig. Input 24V, 3ms]
//       Term 1089 (EL1809) [EL1809 16Ch. Dig. Input 24V, 3ms]
//       Term 1090 (EL1809) [EL1809 16Ch. Dig. Input 24V, 3ms]
//       Term 1091 (EL1809) [EL1809 16Ch. Dig. Input 24V, 3ms]
//       Term 1092 (EL1809) [EL1809 16Ch. Dig. Input 24V, 3ms]
//       Term 1093 (EL1809) [EL1809 16Ch. Dig. Input 24V, 3ms]
//       Term 1094 (EL1809) [EL1809 16Ch. Dig. Input 24V, 3ms]
//       Term 1095 (EL1809) [EL1809 16Ch. Dig. Input 24V, 3ms]
//       Term 1096 (EL1809) [EL1809 16Ch. Dig. Input 24V, 3ms]
//       Term 1097 (EL1809) [EL1809 16Ch. Dig. Input 24V, 3ms]
//       Term 1098 (EL1809) [EL1809 16Ch. Dig. Input 24V, 3ms]
//       Term 1099 (EL1809) [EL1809 16Ch. Dig. Input 24V, 3ms]
//       Term 1100 (EL1809) [EL1809 16Ch. Dig. Input 24V, 3ms]
//       Term 1101 (EL1809) [EL1809 16Ch. Dig. Input 24V, 3ms]
//       Term 1102 (EL1809) [EL1809 16Ch. Dig. Input 24V, 3ms]
//       Term 1103 (EL1809) [EL1809 16Ch. Dig. Input 24V, 3ms]
//       Term 1104 (EL1809) [EL1809 16Ch. Dig. Input 24V, 3ms]
//       Term 1105 (EL1809) [EL1809 16Ch. Dig. Input 24V, 3ms]
//       Term 1106 (EL1809) [EL1809 16Ch. Dig. Input 24V, 3ms]
//       Term 1107 (EL1809) [EL1809 16Ch. Dig. Input 24V, 3ms]
//       Term 1108 (EL1809) [EL1809 16Ch. Dig. Input 24V, 3ms]
//       Term 1109 (EL1809) [EL1809 16Ch. Dig. Input 24V, 3ms]
//       Term 1110 (EL1809) [EL1809 16Ch. Dig. Input 24V, 3ms]
//       Term 1111 (EL1809) [EL1809 16Ch. Dig. Input 24V, 3ms]
//       Term 1112 (EL1809) [EL1809 16Ch. Dig. Input 24V, 3ms]
//       Term 1113 (EL1809) [EL1809 16Ch. Dig. Input 24V, 3ms]
//       Term 1114 (EL1809) [EL1809 16Ch. Dig. Input 24V, 3ms]
//       Term 1115 (EL1809) [EL1809 16Ch. Dig. Input 24V, 3ms]
//       Term 1116 (EL1809) [EL1809 16Ch. Dig. Input 24V, 3ms]
//       Term 1117 (EL1809) [EL1809 16Ch. Dig. Input 24V, 3ms]
//       Term 1118 (EL1809) [EL1809 16Ch. Dig. Input 24V, 3ms]
//       Term 1119 (EL1809) [EL1809 16Ch. Dig. Input 24V, 3ms]
//       Term 1120 (EL1809) [EL1809 16Ch. Dig. Input 24V, 3ms]
//       Term 1121 (EL1809) [EL1809 16Ch. Dig. Input 24V, 3ms]
//       Term 1122 (EL1809) [EL1809 16Ch. Dig. Input 24V, 3ms]
//       Term 1123 (EL1809) [EL1809 16Ch. Dig. Input 24V, 3ms]
//       Term 1124 (EL1809) [EL1809 16Ch. Dig. Input 24V, 3ms]
//       Term 1125 (EL1809) [EL1809 16Ch. Dig. Input 24V, 3ms]
//       Term 1126 (EL1809) [EL1809 16Ch. Dig. Input 24V, 3ms]
//       Term 1127 (EL1809) [EL1809 16Ch. Dig. Input 24V, 3ms]
//       Term 1128 (EL1809) [EL1809 16Ch. Dig. Input 24V, 3ms]
//       Term 1129 (EL1809) [EL1809 16Ch. Dig. Input 24V, 3ms]
//       Term 1130 (EL1809) [EL1809 16Ch. Dig. Input 24V, 3ms]
//       Term 1131 (EL1809) [EL1809 16Ch. Dig. Input 24V, 3ms]
//       Term 1132 (EL1809) [EL1809 16Ch. Dig. Input 24V, 3ms]
//       Term 1134 (EL1809) [EL1809 16Ch. Dig. Input 24V, 3ms]
//       Term 1135 (EL1809) [EL1809 16Ch. Dig. Input 24V, 3ms]
//       Term 1136 (EL1809) [EL1809 16Ch. Dig. Input 24V, 3ms]
//       Term 1137 (EL1809) [EL1809 16Ch. Dig. Input 24V, 3ms]
//       Term 1138 (EL1809) [EL1809 16Ch. Dig. Input 24V, 3ms]
//       Term 1139 (EL1809) [EL1809 16Ch. Dig. Input 24V, 3ms]
//       Term 1140 (EL1809) [EL1809 16Ch. Dig. Input 24V, 3ms]
//       Term 1141 (EL1809) [EL1809 16Ch. Dig. Input 24V, 3ms]
//       Term 1142 (EL1809) [EL1809 16Ch. Dig. Input 24V, 3ms]
//       Term 1143 (EL1809) [EL1809 16Ch. Dig. Input 24V, 3ms]
//       Term 1144 (EL1809) [EL1809 16Ch. Dig. Input 24V, 3ms]
//       Term 1145 (EL1809) [EL1809 16Ch. Dig. Input 24V, 3ms]
//       Term 1146 (EL1809) [EL1809 16Ch. Dig. Input 24V, 3ms]
//       Term 1147 (EL1809) [EL1809 16Ch. Dig. Input 24V, 3ms]
//       Term 1148 (EL1809) [EL1809 16Ch. Dig. Input 24V, 3ms]
//       Term 1149 (EL1809) [EL1809 16Ch. Dig. Input 24V, 3ms]
//       Term 1150 (EL1809) [EL1809 16Ch. Dig. Input 24V, 3ms]
//       Term 1151 (EL1809) [EL1809 16Ch. Dig. Input 24V, 3ms]
//       Term 1154 (EL1809) [EL1809 16Ch. Dig. Input 24V, 3ms]
//       Term 1155 (EL1809) [EL1809 16Ch. Dig. Input 24V, 3ms]
//       Term 1156 (EL1809) [EL1809 16Ch. Dig. Input 24V, 3ms]
//       Term 1157 (EK1110) [EK1110 EtherCAT extension]
// variable links:
//   TcoIoTests/TcoIoTests Instance <-> Device 1 (EtherCAT)
//     PlcTask Inputs/GVL_iXlinker.Device_1_EtherCAT.InfoData.AmsNetId <-> InfoData/AmsNetId
//     PlcTask Inputs/GVL_iXlinker.Device_1_EtherCAT.InfoData.CfgSlaveCount <-> InfoData/CfgSlaveCount
//     PlcTask Inputs/GVL_iXlinker.Device_1_EtherCAT.InfoData.ChangeCount <-> InfoData/ChangeCount
//     PlcTask Inputs/GVL_iXlinker.Device_1_EtherCAT.InfoData.DcToExtTimeOffset <-> InfoData/DcToExtTimeOffset
//     PlcTask Inputs/GVL_iXlinker.Device_1_EtherCAT.InfoData.DcToTcTimeOffset <-> InfoData/DcToTcTimeOffset
//     PlcTask Inputs/GVL_iXlinker.Device_1_EtherCAT.InfoData.DevId <-> InfoData/DevId
//     PlcTask Inputs/GVL_iXlinker.Device_1_EtherCAT.Inputs.DevState <-> Inputs/DevState
//     PlcTask Inputs/GVL_iXlinker.Device_1_EtherCAT.Inputs.Frm0InputToggle <-> Inputs/Frm0InputToggle
//     PlcTask Inputs/GVL_iXlinker.Device_1_EtherCAT.Inputs.Frm0State <-> Inputs/Frm0State
//     PlcTask Inputs/GVL_iXlinker.Device_1_EtherCAT.Inputs.Frm0WcState <-> Inputs/Frm0WcState
//     PlcTask Inputs/GVL_iXlinker.Device_1_EtherCAT.Inputs.SlaveCount <-> Inputs/SlaveCount
//     PlcTask Outputs/GVL_iXlinker.Device_1_EtherCAT.Outputs.DevCtrl <-> Outputs/DevCtrl
//     PlcTask Outputs/GVL_iXlinker.Device_1_EtherCAT.Outputs.Frm0Ctrl <-> Outputs/Frm0Ctrl
//     PlcTask Outputs/GVL_iXlinker.Device_1_EtherCAT.Outputs.Frm0WcCtrl <-> Outputs/Frm0WcCtrl
//   TcoIoTests/TcoIoTests Instance <-> Device 1 (EtherCAT)/Term 1 (EK1200)/Term 2 (EL6002)
//     PlcTask Inputs/GVL_iXlinker.Device_1_EtherCAT.Term_1_EK1200.Term_2_EL6002.COM_TxPDO_Map_Inputs_Channel_1.Data_In[0] <-> COM TxPDO-Map Inputs Channel 1/Data In 0
//     PlcTask Inputs/GVL_iXlinker.Device_1_EtherCAT.Term_1_EK1200.Term_2_EL6002.COM_TxPDO_Map_Inputs_Channel_1.Data_In[10] <-> COM TxPDO-Map Inputs Channel 1/Data In 10
//     PlcTask Inputs/GVL_iXlinker.Device_1_EtherCAT.Term_1_EK1200.Term_2_EL6002.COM_TxPDO_Map_Inputs_Channel_1.Data_In[11] <-> COM TxPDO-Map Inputs Channel 1/Data In 11
//     PlcTask Inputs/GVL_iXlinker.Device_1_EtherCAT.Term_1_EK1200.Term_2_EL6002.COM_TxPDO_Map_Inputs_Channel_1.Data_In[12] <-> COM TxPDO-Map Inputs Channel 1/Data In 12
//     PlcTask Inputs/GVL_iXlinker.Device_1_EtherCAT.Term_1_EK1200.Term_2_EL6002.COM_TxPDO_Map_Inputs_Channel_1.Data_In[13] <-> COM TxPDO-Map Inputs Channel 1/Data In 13
//     PlcTask Inputs/GVL_iXlinker.Device_1_EtherCAT.Term_1_EK1200.Term_2_EL6002.COM_TxPDO_Map_Inputs_Channel_1.Data_In[14] <-> COM TxPDO-Map Inputs Channel 1/Data In 14
//     PlcTask Inputs/GVL_iXlinker.Device_1_EtherCAT.Term_1_EK1200.Term_2_EL6002.COM_TxPDO_Map_Inputs_Channel_1.Data_In[15] <-> COM TxPDO-Map Inputs Channel 1/Data In 15
//     PlcTask Inputs/GVL_iXlinker.Device_1_EtherCAT.Term_1_EK1200.Term_2_EL6002.COM_TxPDO_Map_Inputs_Channel_1.Data_In[16] <-> COM TxPDO-Map Inputs Channel 1/Data In 16
//     PlcTask Inputs/GVL_iXlinker.Device_1_EtherCAT.Term_1_EK1200.Term_2_EL6002.COM_TxPDO_Map_Inputs_Channel_1.Data_In[17] <-> COM TxPDO-Map Inputs Channel 1/Data In 17
//     PlcTask Inputs/GVL_iXlinker.Device_1_EtherCAT.Term_1_EK1200.Term_2_EL6002.COM_TxPDO_Map_Inputs_Channel_1.Data_In[18] <-> COM TxPDO-Map Inputs Channel 1/Data In 18
//     PlcTask Inputs/GVL_iXlinker.Device_1_EtherCAT.Term_1_EK1200.Term_2_EL6002.COM_TxPDO_Map_Inputs_Channel_1.Data_In[19] <-> COM TxPDO-Map Inputs Channel 1/Data In 19
//     PlcTask Inputs/GVL_iXlinker.Device_1_EtherCAT.Term_1_EK1200.Term_2_EL6002.COM_TxPDO_Map_Inputs_Channel_1.Data_In[1] <-> COM TxPDO-Map Inputs Channel 1/Data In 1
//     PlcTask Inputs/GVL_iXlinker.Device_1_EtherCAT.Term_1_EK1200.Term_2_EL6002.COM_TxPDO_Map_Inputs_Channel_1.Data_In[20] <-> COM TxPDO-Map Inputs Channel 1/Data In 20
//     PlcTask Inputs/GVL_iXlinker.Device_1_EtherCAT.Term_1_EK1200.Term_2_EL6002.COM_TxPDO_Map_Inputs_Channel_1.Data_In[21] <-> COM TxPDO-Map Inputs Channel 1/Data In 21
//     PlcTask Inputs/GVL_iXlinker.Device_1_EtherCAT.Term_1_EK1200.Term_2_EL6002.COM_TxPDO_Map_Inputs_Channel_1.Data_In[2] <-> COM TxPDO-Map Inputs Channel 1/Data In 2
//     PlcTask Inputs/GVL_iXlinker.Device_1_EtherCAT.Term_1_EK1200.Term_2_EL6002.COM_TxPDO_Map_Inputs_Channel_1.Data_In[3] <-> COM TxPDO-Map Inputs Channel 1/Data In 3
//     PlcTask Inputs/GVL_iXlinker.Device_1_EtherCAT.Term_1_EK1200.Term_2_EL6002.COM_TxPDO_Map_Inputs_Channel_1.Data_In[4] <-> COM TxPDO-Map Inputs Channel 1/Data In 4
//     PlcTask Inputs/GVL_iXlinker.Device_1_EtherCAT.Term_1_EK1200.Term_2_EL6002.COM_TxPDO_Map_Inputs_Channel_1.Data_In[5] <-> COM TxPDO-Map Inputs Channel 1/Data In 5
//     PlcTask Inputs/GVL_iXlinker.Device_1_EtherCAT.Term_1_EK1200.Term_2_EL6002.COM_TxPDO_Map_Inputs_Channel_1.Data_In[6] <-> COM TxPDO-Map Inputs Channel 1/Data In 6
//     PlcTask Inputs/GVL_iXlinker.Device_1_EtherCAT.Term_1_EK1200.Term_2_EL6002.COM_TxPDO_Map_Inputs_Channel_1.Data_In[7] <-> COM TxPDO-Map Inputs Channel 1/Data In 7
//     PlcTask Inputs/GVL_iXlinker.Device_1_EtherCAT.Term_1_EK1200.Term_2_EL6002.COM_TxPDO_Map_Inputs_Channel_1.Data_In[8] <-> COM TxPDO-Map Inputs Channel 1/Data In 8
//     PlcTask Inputs/GVL_iXlinker.Device_1_EtherCAT.Term_1_EK1200.Term_2_EL6002.COM_TxPDO_Map_Inputs_Channel_1.Data_In[9] <-> COM TxPDO-Map Inputs Channel 1/Data In 9
//     PlcTask Inputs/GVL_iXlinker.Device_1_EtherCAT.Term_1_EK1200.Term_2_EL6002.COM_TxPDO_Map_Inputs_Channel_2.Data_In[0] <-> COM TxPDO-Map Inputs Channel 2/Data In 0
//     PlcTask Inputs/GVL_iXlinker.Device_1_EtherCAT.Term_1_EK1200.Term_2_EL6002.COM_TxPDO_Map_Inputs_Channel_2.Data_In[10] <-> COM TxPDO-Map Inputs Channel 2/Data In 10
//     PlcTask Inputs/GVL_iXlinker.Device_1_EtherCAT.Term_1_EK1200.Term_2_EL6002.COM_TxPDO_Map_Inputs_Channel_2.Data_In[11] <-> COM TxPDO-Map Inputs Channel 2/Data In 11
//     PlcTask Inputs/GVL_iXlinker.Device_1_EtherCAT.Term_1_EK1200.Term_2_EL6002.COM_TxPDO_Map_Inputs_Channel_2.Data_In[12] <-> COM TxPDO-Map Inputs Channel 2/Data In 12
//     PlcTask Inputs/GVL_iXlinker.Device_1_EtherCAT.Term_1_EK1200.Term_2_EL6002.COM_TxPDO_Map_Inputs_Channel_2.Data_In[13] <-> COM TxPDO-Map Inputs Channel 2/Data In 13
//     PlcTask Inputs/GVL_iXlinker.Device_1_EtherCAT.Term_1_EK1200.Term_2_EL6002.COM_TxPDO_Map_Inputs_Channel_2.Data_In[14] <-> COM TxPDO-Map Inputs Channel 2/Data In 14
//     PlcTask Inputs/GVL_iXlinker.Device_1_EtherCAT.Term_1_EK1200.Term_2_EL6002.COM_TxPDO_Map_Inputs_Channel_2.Data_In[15] <-> COM TxPDO-Map Inputs Channel 2/Data In 15
//     PlcTask Inputs/GVL_iXlinker.Device_1_EtherCAT.Term_1_EK1200.Term_2_EL6002.COM_TxPDO_Map_Inputs_Channel_2.Data_In[16] <-> COM TxPDO-Map Inputs Channel 2/Data In 16
//     PlcTask Inputs/GVL_iXlinker.Device_1_EtherCAT.Term_1_EK1200.Term_2_EL6002.COM_TxPDO_Map_Inputs_Channel_2.Data_In[17] <-> COM TxPDO-Map Inputs Channel 2/Data In 17
//     PlcTask Inputs/GVL_iXlinker.Device_1_EtherCAT.Term_1_EK1200.Term_2_EL6002.COM_TxPDO_Map_Inputs_Channel_2.Data_In[18] <-> COM TxPDO-Map Inputs Channel 2/Data In 18
//     PlcTask Inputs/GVL_iXlinker.Device_1_EtherCAT.Term_1_EK1200.Term_2_EL6002.COM_TxPDO_Map_Inputs_Channel_2.Data_In[19] <-> COM TxPDO-Map Inputs Channel 2/Data In 19
//     PlcTask Inputs/GVL_iXlinker.Device_1_EtherCAT.Term_1_EK1200.Term_2_EL6002.COM_TxPDO_Map_Inputs_Channel_2.Data_In[1] <-> COM TxPDO-Map Inputs Channel 2/Data In 1
//     PlcTask Inputs/GVL_iXlinker.Device_1_EtherCAT.Term_1_EK1200.Term_2_EL6002.COM_TxPDO_Map_Inputs_Channel_2.Data_In[20] <-> COM TxPDO-Map Inputs Channel 2/Data In 20
//     PlcTask Inputs/GVL_iXlinker.Device_1_EtherCAT.Term_1_EK1200.Term_2_EL6002.COM_TxPDO_Map_Inputs_Channel_2.Data_In[21] <-> COM TxPDO-Map Inputs Channel 2/Data In 21
//     PlcTask Inputs/GVL_iXlinker.Device_1_EtherCAT.Term_1_EK1200.Term_2_EL6002.COM_TxPDO_Map_Inputs_Channel_2.Data_In[2] <-> COM TxPDO-Map Inputs Channel 2/Data In 2
//     PlcTask Inputs/GVL_iXlinker.Device_1_EtherCAT.Term_1_EK1200.Term_2_EL6002.COM_TxPDO_Map_Inputs_Channel_2.Data_In[3] <-> COM TxPDO-Map Inputs Channel 2/Data In 3
//     PlcTask Inputs/GVL_iXlinker.Device_1_EtherCAT.Term_1_EK1200.Term_2_EL6002.COM_TxPDO_Map_Inputs_Channel_2.Data_In[4] <-> COM TxPDO-Map Inputs Channel 2/Data In 4
//     PlcTask Inputs/GVL_iXlinker.Device_1_EtherCAT.Term_1_EK1200.Term_2_EL6002.COM_TxPDO_Map_Inputs_Channel_2.Data_In[5] <-> COM TxPDO-Map Inputs Channel 2/Data In 5
//     PlcTask Inputs/GVL_iXlinker.Device_1_EtherCAT.Term_1_EK1200.Term_2_EL6002.COM_TxPDO_Map_Inputs_Channel_2.Data_In[6] <-> COM TxPDO-Map Inputs Channel 2/Data In 6
//     PlcTask Inputs/GVL_iXlinker.Device_1_EtherCAT.Term_1_EK1200.Term_2_EL6002.COM_TxPDO_Map_Inputs_Channel_2.Data_In[7] <-> COM TxPDO-Map Inputs Channel 2/Data In 7
//     PlcTask Inputs/GVL_iXlinker.Device_1_EtherCAT.Term_1_EK1200.Term_2_EL6002.COM_TxPDO_Map_Inputs_Channel_2.Data_In[8] <-> COM TxPDO-Map Inputs Channel 2/Data In 8
//     PlcTask Inputs/GVL_iXlinker.Device_1_EtherCAT.Term_1_EK1200.Term_2_EL6002.COM_TxPDO_Map_Inputs_Channel_2.Data_In[9] <-> COM TxPDO-Map Inputs Channel 2/Data In 9
//     PlcTask Inputs/GVL_iXlinker.Device_1_EtherCAT.Term_1_EK1200.Term_2_EL6002.COM_TxPDO_Map_Inputs_Channel_1.Status/Buffer_full <-> COM TxPDO-Map Inputs Channel 1/Status/Buffer full
//     PlcTask Inputs/GVL_iXlinker.Device_1_EtherCAT.Term_1_EK1200.Term_2_EL6002.COM_TxPDO_Map_Inputs_Channel_2.Status/Buffer_full <-> COM TxPDO-Map Inputs Channel 2/Status/Buffer full
//     PlcTask Inputs/GVL_iXlinker.Device_1_EtherCAT.Term_1_EK1200.Term_2_EL6002.COM_TxPDO_Map_Inputs_Channel_1.Status/Framing_error <-> COM TxPDO-Map Inputs Channel 1/Status/Framing error
//     PlcTask Inputs/GVL_iXlinker.Device_1_EtherCAT.Term_1_EK1200.Term_2_EL6002.COM_TxPDO_Map_Inputs_Channel_2.Status/Framing_error <-> COM TxPDO-Map Inputs Channel 2/Status/Framing error
//     PlcTask Inputs/GVL_iXlinker.Device_1_EtherCAT.Term_1_EK1200.Term_2_EL6002.COM_TxPDO_Map_Inputs_Channel_1.Status/Init_accepted <-> COM TxPDO-Map Inputs Channel 1/Status/Init accepted
//     PlcTask Inputs/GVL_iXlinker.Device_1_EtherCAT.Term_1_EK1200.Term_2_EL6002.COM_TxPDO_Map_Inputs_Channel_2.Status/Init_accepted <-> COM TxPDO-Map Inputs Channel 2/Status/Init accepted
//     PlcTask Inputs/GVL_iXlinker.Device_1_EtherCAT.Term_1_EK1200.Term_2_EL6002.COM_TxPDO_Map_Inputs_Channel_1.Status/Input_length <-> COM TxPDO-Map Inputs Channel 1/Status/Input length
//     PlcTask Inputs/GVL_iXlinker.Device_1_EtherCAT.Term_1_EK1200.Term_2_EL6002.COM_TxPDO_Map_Inputs_Channel_2.Status/Input_length <-> COM TxPDO-Map Inputs Channel 2/Status/Input length
//     PlcTask Inputs/GVL_iXlinker.Device_1_EtherCAT.Term_1_EK1200.Term_2_EL6002.COM_TxPDO_Map_Inputs_Channel_1.Status/Overrun_error <-> COM TxPDO-Map Inputs Channel 1/Status/Overrun error
//     PlcTask Inputs/GVL_iXlinker.Device_1_EtherCAT.Term_1_EK1200.Term_2_EL6002.COM_TxPDO_Map_Inputs_Channel_2.Status/Overrun_error <-> COM TxPDO-Map Inputs Channel 2/Status/Overrun error
//     PlcTask Inputs/GVL_iXlinker.Device_1_EtherCAT.Term_1_EK1200.Term_2_EL6002.COM_TxPDO_Map_Inputs_Channel_1.Status/Parity_error <-> COM TxPDO-Map Inputs Channel 1/Status/Parity error
//     PlcTask Inputs/GVL_iXlinker.Device_1_EtherCAT.Term_1_EK1200.Term_2_EL6002.COM_TxPDO_Map_Inputs_Channel_2.Status/Parity_error <-> COM TxPDO-Map Inputs Channel 2/Status/Parity error
//     PlcTask Inputs/GVL_iXlinker.Device_1_EtherCAT.Term_1_EK1200.Term_2_EL6002.COM_TxPDO_Map_Inputs_Channel_1.Status/Receive_request <-> COM TxPDO-Map Inputs Channel 1/Status/Receive request
//     PlcTask Inputs/GVL_iXlinker.Device_1_EtherCAT.Term_1_EK1200.Term_2_EL6002.COM_TxPDO_Map_Inputs_Channel_2.Status/Receive_request <-> COM TxPDO-Map Inputs Channel 2/Status/Receive request
//     PlcTask Inputs/GVL_iXlinker.Device_1_EtherCAT.Term_1_EK1200.Term_2_EL6002.COM_TxPDO_Map_Inputs_Channel_1.Status/Transmit_accepted <-> COM TxPDO-Map Inputs Channel 1/Status/Transmit accepted
//     PlcTask Inputs/GVL_iXlinker.Device_1_EtherCAT.Term_1_EK1200.Term_2_EL6002.COM_TxPDO_Map_Inputs_Channel_2.Status/Transmit_accepted <-> COM TxPDO-Map Inputs Channel 2/Status/Transmit accepted
//     PlcTask Inputs/GVL_iXlinker.Device_1_EtherCAT.Term_1_EK1200.Term_2_EL6002.InfoData.AdsAddr <-> InfoData/AdsAddr
//     PlcTask Inputs/GVL_iXlinker.Device_1_EtherCAT.Term_1_EK1200.Term_2_EL6002.InfoData.State <-> InfoData/State
//     PlcTask Inputs/GVL_iXlinker.Device_1_EtherCAT.Term_1_EK1200.Term_2_EL6002.WcState.InputToggle <-> WcState/InputToggle
//     PlcTask Inputs/GVL_iXlinker.Device_1_EtherCAT.Term_1_EK1200.Term_2_EL6002.WcState.WcState <-> WcState/WcState
//     PlcTask Outputs/GVL_iXlinker.Device_1_EtherCAT.Term_1_EK1200.Term_2_EL6002.COM_RxPDO_Map_Outputs_Channel_1.Ctrl/Init_request <-> COM RxPDO-Map Outputs Channel 1/Ctrl/Init request
//     PlcTask Outputs/GVL_iXlinker.Device_1_EtherCAT.Term_1_EK1200.Term_2_EL6002.COM_RxPDO_Map_Outputs_Channel_2.Ctrl/Init_request <-> COM RxPDO-Map Outputs Channel 2/Ctrl/Init request
//     PlcTask Outputs/GVL_iXlinker.Device_1_EtherCAT.Term_1_EK1200.Term_2_EL6002.COM_RxPDO_Map_Outputs_Channel_1.Ctrl/Output_length <-> COM RxPDO-Map Outputs Channel 1/Ctrl/Output length
//     PlcTask Outputs/GVL_iXlinker.Device_1_EtherCAT.Term_1_EK1200.Term_2_EL6002.COM_RxPDO_Map_Outputs_Channel_2.Ctrl/Output_length <-> COM RxPDO-Map Outputs Channel 2/Ctrl/Output length
//     PlcTask Outputs/GVL_iXlinker.Device_1_EtherCAT.Term_1_EK1200.Term_2_EL6002.COM_RxPDO_Map_Outputs_Channel_1.Ctrl/Receive_accepted <-> COM RxPDO-Map Outputs Channel 1/Ctrl/Receive accepted
//     PlcTask Outputs/GVL_iXlinker.Device_1_EtherCAT.Term_1_EK1200.Term_2_EL6002.COM_RxPDO_Map_Outputs_Channel_2.Ctrl/Receive_accepted <-> COM RxPDO-Map Outputs Channel 2/Ctrl/Receive accepted
//     PlcTask Outputs/GVL_iXlinker.Device_1_EtherCAT.Term_1_EK1200.Term_2_EL6002.COM_RxPDO_Map_Outputs_Channel_1.Ctrl/Send_continuous <-> COM RxPDO-Map Outputs Channel 1/Ctrl/Send continuous
//     PlcTask Outputs/GVL_iXlinker.Device_1_EtherCAT.Term_1_EK1200.Term_2_EL6002.COM_RxPDO_Map_Outputs_Channel_2.Ctrl/Send_continuous <-> COM RxPDO-Map Outputs Channel 2/Ctrl/Send continuous
//     PlcTask Outputs/GVL_iXlinker.Device_1_EtherCAT.Term_1_EK1200.Term_2_EL6002.COM_RxPDO_Map_Outputs_Channel_1.Ctrl/Transmit_request <-> COM RxPDO-Map Outputs Channel 1/Ctrl/Transmit request
//     PlcTask Outputs/GVL_iXlinker.Device_1_EtherCAT.Term_1_EK1200.Term_2_EL6002.COM_RxPDO_Map_Outputs_Channel_2.Ctrl/Transmit_request <-> COM RxPDO-Map Outputs Channel 2/Ctrl/Transmit request
//     PlcTask Outputs/GVL_iXlinker.Device_1_EtherCAT.Term_1_EK1200.Term_2_EL6002.COM_RxPDO_Map_Outputs_Channel_1.Data_Out[0] <-> COM RxPDO-Map Outputs Channel 1/Data Out 0
//     PlcTask Outputs/GVL_iXlinker.Device_1_EtherCAT.Term_1_EK1200.Term_2_EL6002.COM_RxPDO_Map_Outputs_Channel_1.Data_Out[10] <-> COM RxPDO-Map Outputs Channel 1/Data Out 10
//     PlcTask Outputs/GVL_iXlinker.Device_1_EtherCAT.Term_1_EK1200.Term_2_EL6002.COM_RxPDO_Map_Outputs_Channel_1.Data_Out[11] <-> COM RxPDO-Map Outputs Channel 1/Data Out 11
//     PlcTask Outputs/GVL_iXlinker.Device_1_EtherCAT.Term_1_EK1200.Term_2_EL6002.COM_RxPDO_Map_Outputs_Channel_1.Data_Out[12] <-> COM RxPDO-Map Outputs Channel 1/Data Out 12
//     PlcTask Outputs/GVL_iXlinker.Device_1_EtherCAT.Term_1_EK1200.Term_2_EL6002.COM_RxPDO_Map_Outputs_Channel_1.Data_Out[13] <-> COM RxPDO-Map Outputs Channel 1/Data Out 13
//     PlcTask Outputs/GVL_iXlinker.Device_1_EtherCAT.Term_1_EK1200.Term_2_EL6002.COM_RxPDO_Map_Outputs_Channel_1.Data_Out[14] <-> COM RxPDO-Map Outputs Channel 1/Data Out 14
//     PlcTask Outputs/GVL_iXlinker.Device_1_EtherCAT.Term_1_EK1200.Term_2_EL6002.COM_RxPDO_Map_Outputs_Channel_1.Data_Out[15] <-> COM RxPDO-Map Outputs Channel 1/Data Out 15
//     PlcTask Outputs/GVL_iXlinker.Device_1_EtherCAT.Term_1_EK1200.Term_2_EL6002.COM_RxPDO_Map_Outputs_Channel_1.Data_Out[16] <-> COM RxPDO-Map Outputs Channel 1/Data Out 16
//     PlcTask Outputs/GVL_iXlinker.Device_1_EtherCAT.Term_1_EK1200.Term_2_EL6002.COM_RxPDO_Map_Outputs_Channel_1.Data_Out[17] <-> COM RxPDO-Map Outputs Channel 1/Data Out 17
//     PlcTask Outputs/GVL_iXlinker.Device_1_EtherCAT.Term_1_EK1200.Term_2_EL6002.COM_RxPDO_Map_Outputs_Channel_1.Data_Out[18] <-> COM RxPDO-Map Outputs Channel 1/Data Out 18
//     PlcTask Outputs/GVL_iXlinker.Device_1_EtherCAT.Term_1_EK1200.Term_2_EL6002.COM_RxPDO_Map_Outputs_Channel_1.Data_Out[19] <-> COM RxPDO-Map Outputs Channel 1/Data Out 19
//     PlcTask Outputs/GVL_iXlinker.Device_1_EtherCAT.Term_1_EK1200.Term_2_EL6002.COM_RxPDO_Map_Outputs_Channel_1.Data_Out[1] <-> COM RxPDO-Map Outputs Channel 1/Data Out 1
//     PlcTask Outputs/GVL_iXlinker.Device_1_EtherCAT.Term_1_EK1200.Term_2_EL6002.COM_RxPDO_Map_Outputs_Channel_1.Data_Out[20] <-> COM RxPDO-Map Outputs Channel 1/Data Out 20
//     PlcTask Outputs/GVL_iXlinker.Device_1_EtherCAT.Term_1_EK1200.Term_2_EL6002.COM_RxPDO_Map_Outputs_Channel_1.Data_Out[21] <-> COM RxPDO-Map Outputs Channel 1/Data Out 21
//     PlcTask Outputs/GVL_iXlinker.Device_1_EtherCAT.Term_1_EK1200.Term_2_EL6002.COM_RxPDO_Map_Outputs_Channel_1.Data_Out[2] <-> COM RxPDO-Map Outputs Channel 1/Data Out 2
